screen "C5_GraphicView_2" 1024x768, template "T_C05"
   GraphicView "PNG_160x60_FitF" at 6,40 size 160x60; Picture "G_PNG"
   TextField "Label_PNG_160x60_FitF" at 6,102 size 113x20; Text 'PNG_160x60_FitF'
   GraphicView "PNG_160x60_FitT" at 182,40 size 160x60; Picture "G_PNG"
   TextField "Label_PNG_160x60_FitT" at 182,102 size 114x20; Text 'PNG_160x60_FitT'
   GraphicView "PNG_60x120_FitF" at 358,40 size 60x120; Picture "G_PNG"
   TextField "Label_PNG_60x120_FitF" at 358,162 size 113x20; Text 'PNG_60x120_FitF'
   GraphicView "PNG_60x120_FitT" at 534,40 size 60x120; Picture "G_PNG"
   TextField "Label_PNG_60x120_FitT" at 534,162 size 114x20; Text 'PNG_60x120_FitT'
   GraphicView "PNG_80x80_FitF" at 710,40 size 80x80; Picture "G_PNG"
   TextField "Label_PNG_80x80_FitF" at 710,122 size 105x20; Text 'PNG_80x80_FitF'
   GraphicView "PNG_80x80_FitT" at 6,182 size 80x80; Picture "G_PNG"
   TextField "Label_PNG_80x80_FitT" at 6,264 size 106x20; Text 'PNG_80x80_FitT'
   GraphicView "TALL_160x60_FitF" at 182,182 size 160x60; Picture "G_TALL"
   TextField "Label_TALL_160x60_FitF" at 182,244 size 120x20; Text 'TALL_160x60_FitF'
   GraphicView "TALL_160x60_FitT" at 358,182 size 160x60; Picture "G_TALL"
   TextField "Label_TALL_160x60_FitT" at 358,244 size 121x20; Text 'TALL_160x60_FitT'
   GraphicView "TALL_60x120_FitF" at 534,182 size 60x120; Picture "G_TALL"
   TextField "Label_TALL_60x120_FitF" at 534,304 size 120x20; Text 'TALL_60x120_FitF'
   GraphicView "TALL_60x120_FitT" at 710,182 size 60x120; Picture "G_TALL"
   TextField "Label_TALL_60x120_FitT" at 710,304 size 121x20; Text 'TALL_60x120_FitT'
   GraphicView "TALL_80x80_FitF" at 6,324 size 80x80; Picture "G_TALL"
   TextField "Label_TALL_80x80_FitF" at 6,406 size 112x20; Text 'TALL_80x80_FitF'
   GraphicView "TALL_80x80_FitT" at 182,324 size 80x80; Picture "G_TALL"
   TextField "Label_TALL_80x80_FitT" at 182,406 size 113x20; Text 'TALL_80x80_FitT'
   GraphicView "WIDE_160x60_FitF" at 358,324 size 160x60; Picture "G_WIDE"
   TextField "Label_WIDE_160x60_FitF" at 358,386 size 123x20; Text 'WIDE_160x60_FitF'
   GraphicView "WIDE_160x60_FitT" at 534,324 size 160x60; Picture "G_WIDE"
   TextField "Label_WIDE_160x60_FitT" at 534,386 size 124x20; Text 'WIDE_160x60_FitT'
   GraphicView "WIDE_60x120_FitF" at 710,324 size 60x120; Picture "G_WIDE"
   TextField "Label_WIDE_60x120_FitF" at 710,446 size 123x20; Text 'WIDE_60x120_FitF'
   GraphicView "WIDE_60x120_FitT" at 6,466 size 60x120; Picture "G_WIDE"
   TextField "Label_WIDE_60x120_FitT" at 6,588 size 124x20; Text 'WIDE_60x120_FitT'
   GraphicView "WIDE_80x80_FitF" at 182,466 size 80x80; Picture "G_WIDE"
   TextField "Label_WIDE_80x80_FitF" at 182,548 size 115x20; Text 'WIDE_80x80_FitF'
   GraphicView "WIDE_80x80_FitT" at 358,466 size 80x80; Picture "G_WIDE"
   TextField "Label_WIDE_80x80_FitT" at 358,548 size 116x20; Text 'WIDE_80x80_FitT'
   GraphicView "BMP_Transparent" at 534,466 size 120x80; Picture "G_BMP"
   TextField "Label_BMP_Transparent" at 534,548 size 120x20; Text 'BMP_Transparent'
   GraphicView "PNG_BackTransparent" at 710,466 size 120x80; Picture "G_PNG"
   TextField "Label_PNG_BackTransparent" at 710,548 size 147x20; Text 'PNG_BackTransparent'
   IOField "State" at 4,742 size 60x22; FormatPattern 9
      ProcessValue <- "D_State"
   Button "S1" at 70,742 size 40x22; TextOff 'S1'
      on Click: "SetS1"()
   Button "S2" at 114,742 size 40x22; TextOff 'S2'
      on Click: "SetS2"()
   Button "S3" at 158,742 size 40x22; TextOff 'S3'
      on Click: "SetS3"()
   Button "S4" at 202,742 size 40x22; TextOff 'S4'
      on Click: "SetS4"()
   Button "Next" at 980,742 size 40x22; TextOff 'Next'
      on Click: ActivateScreen("C5_Lists", 0)

screen "C5_Lists" 1024x768, template "T_C05"
   SymbolicIOField "SIO_TL_Value" at 6,40 size 160x30; TextOff '0'; TextOn '1'; TextList "TL_Value"
      ProcessValue <- "D_TL"
   TextField "Label_SIO_TL_Value" at 6,72 size 93x20; Text 'SIO_TL_Value'
   SymbolicIOField "SIO_TL_Bit" at 182,40 size 160x30; TextOff '0'; TextOn '1'; TextList "TL_Bit"
      ProcessValue <- "D_Bool"
   TextField "Label_SIO_TL_Bit" at 182,72 size 74x20; Text 'SIO_TL_Bit'
   SymbolicIOField "SIO_TL_BitNo" at 358,40 size 160x30; TextOff '0'; TextOn '1'; TextList "TL_BitNo"
      ProcessValue <- "D_Bits"
   TextField "Label_SIO_TL_BitNo" at 358,72 size 90x20; Text 'SIO_TL_BitNo'
   SymbolicIOField "SIO_TL_Value_Out" at 534,40 size 160x30; TextOff '0'; TextOn '1'; TextList "TL_Value"
      ProcessValue <- "D_TL"
   TextField "Label_SIO_TL_Value_Out" at 534,72 size 124x20; Text 'SIO_TL_Value_Out'
   GraphicIOField "GIO_GL_Value" at 710,40 size 120x80; PictureList "GL_Value"
      ProcessValue <- "D_TL"
   TextField "Label_GIO_GL_Value" at 710,122 size 94x20; Text 'GIO_GL_Value'
   GraphicIOField "GIO_GL_Bit" at 6,142 size 120x80; PictureList "GL_Bit"
      ProcessValue <- "D_Bool"
   TextField "Label_GIO_GL_Bit" at 6,224 size 75x20; Text 'GIO_GL_Bit'
   GraphicIOField "GIO_GL_BitNo" at 182,142 size 120x80; PictureList "GL_BitNo"
      ProcessValue <- "D_Bits"
   TextField "Label_GIO_GL_BitNo" at 182,224 size 91x20; Text 'GIO_GL_BitNo'
   GraphicIOField "GIO_GL_Value_Out" at 358,142 size 120x80; PictureList "GL_Value"
      ProcessValue <- "D_TL"
   TextField "Label_GIO_GL_Value_Out" at 358,224 size 125x20; Text 'GIO_GL_Value_Out'
   IOField "State" at 4,742 size 60x22; FormatPattern 9
      ProcessValue <- "D_State"
   Button "S1" at 70,742 size 40x22; TextOff 'S1'
      on Click: "SetS1"()
   Button "S2" at 114,742 size 40x22; TextOff 'S2'
      on Click: "SetS2"()
   Button "S3" at 158,742 size 40x22; TextOff 'S3'
      on Click: "SetS3"()
   Button "S4" at 202,742 size 40x22; TextOff 'S4'
      on Click: "SetS4"()
   Button "Next" at 980,742 size 40x22; TextOff 'Next'
      on Click: ActivateScreen("C5_Buttons", 0)

Template "T_C05" 1024x768
   TextField "T_Title" at 8,6 size 185x21; Text 'Template T_C05 (header)'
   DateTimeField "T_Clock" at 834,4 size 189x26

PopupScreen "Popup_C05" 300x200
   TextField "Pop_Title" at 10,10 size 175x20; Text 'Pop-up screen Popup_C05'
   GraphicView "Pop_Graphic" at 10,40 size 120x80; Picture "G_PNG"
   IOField "Pop_Value" at 150,60 size 120x30; FormatPattern s99999
      ProcessValue <- "D_Int"
   Button "Pop_Close" at 200,160 size 80x22; TextOff 'Close'
      on Click: function_efd93a16("Popup_C05", 200, 120, -1, -1, 1)

screen "C5_Structure" 1024x768, template "T_C05"
   Group "Group_A" at 10,50 size 300x85
   TextField "Label_Group_A (contains Group_B)" at 10,140 size 190x20; Text 'Group_A (contains Group_B)'
   TextField "Layer0_Text" at 352,52 size 54x20; Text 'Layer 0'
   TextField "Label_Layers 0-3 (layer 2 VisibleES false)" at 350,200 size 231x20; Text 'Layers 0-3 (layer 2 VisibleES false)'
   IOField "State" at 4,742 size 60x22; FormatPattern 9
      ProcessValue <- "D_State"
   Button "S1" at 70,742 size 40x22; TextOff 'S1'
      on Click: "SetS1"()
   Button "S2" at 114,742 size 40x22; TextOff 'S2'
      on Click: "SetS2"()
   Button "S3" at 158,742 size 40x22; TextOff 'S3'
      on Click: "SetS3"()
   Button "S4" at 202,742 size 40x22; TextOff 'S4'
      on Click: "SetS4"()
   Button "Popup" at 246,742 size 60x22; TextOff 'Popup'
      on Click: function_efd93a16("Popup_C05", 200, 120, -1, -1, 1)
   Button "SlideIn" at 310,742 size 60x22; TextOff 'Slide'
      on Click: "C5_ToggleSlideIn"()
   Button "Next" at 980,742 size 40x22; TextOff 'Next'
      on Click: ActivateScreen("C5_GraphicView_1", 0)
   Group "Group_B" at 210,50 size 100x85
   TextField "GB_Text" at 210,115 size 59x20; Text 'Group_B'
   TextField "Layer1_Text" at 382,72 size 54x20; Text 'Layer 1'
   TextField "Layer2_Text" at 412,92 size 54x20; Text 'Layer 2'
   TextField "Layer3_Text" at 442,112 size 54x20; Text 'Layer 3'

screen "C6_Faceplates" 1024x768
   ScreenModuleView "FP_Dyn" at 10,10 size 300x150; ScreenModuleType ""; Guid_{11997190-83750} 'Tags D_Int D_Range D_Pct'
      Guid_{11997190-83886} <- "D_Int"
      Guid_{11997190-83896} <- "D_Range"
      Guid_{11997190-83898} <- "D_Pct"
      Guid_{11997190-83900} <- "D_Vis"
   TextField "Label_FP_Dyn" at 10,162 size 52x20; Text 'FP_Dyn'
   ScreenModuleView "FP_Static" at 330,10 size 300x150; ScreenModuleType ""; Guid_{11997190-83750} 'Static values'
   TextField "Label_FP_Static" at 330,162 size 65x20; Text 'FP_Static'
   ScreenModuleView "FP_Alt" at 10,186 size 300x150; ScreenModuleType ""; Guid_{11997190-83750} 'Tags D_SInt D_TL D_UInt'
      Guid_{11997190-83886} <- "D_SInt"
      Guid_{11997190-83896} <- "D_TL"
      Guid_{11997190-83898} <- "D_UInt"
      Guid_{11997190-83900} <- "D_En"
   TextField "Label_FP_Alt" at 10,338 size 46x20; Text 'FP_Alt'
   ScreenModuleView "FP_Move" at 330,186 size 300x150; ScreenModuleType ""; Guid_{11997190-83750} 'Moved by D_Pct'
      Guid_{11997190-83886} <- "D_Int"
      Guid_{11997190-83896} <- "D_Range"
      Guid_{11997190-83898} <- "D_Pct"
      Guid_{11997190-83900} <- "D_Vis"
      HorizontalMovement <- "D_Pct"
   TextField "Label_FP_Move" at 330,338 size 62x20; Text 'FP_Move'
   IOField "State" at 4,742 size 60x22; FormatPattern 9
      ProcessValue <- "D_State"
   Button "S1" at 70,742 size 40x22; TextOff 'S1'
      on Click: "SetS1"()
   Button "S2" at 114,742 size 40x22; TextOff 'S2'
      on Click: "SetS2"()
   Button "S3" at 158,742 size 40x22; TextOff 'S3'
      on Click: "SetS3"()
   Button "S4" at 202,742 size 40x22; TextOff 'S4'
      on Click: "SetS4"()
   Button "Next" at 980,742 size 40x22; TextOff 'Next'
      on Click: ActivateScreen("C6_Faceplates", 0)

VB script "C5_ToggleSlideIn"
   ' slide-in screens are not available on WinCC RT Advanced

VB script "SetS1"
   SmartTags("D_State") = 1
   SmartTags("D_Bool") = False
   SmartTags("D_SInt") = -128
   SmartTags("D_Int") = -32768
   SmartTags("D_DInt") = -2147483648
   SmartTags("D_USInt") = 0
   SmartTags("D_UInt") = 0
   SmartTags("D_UDInt") = 0
   SmartTags("D_Real") = -999.999
   SmartTags("D_LReal") = -0.00000015
   SmartTags("D_String") = ""
   SmartTags("D_DateTime") = DateSerial(1990, 1, 1) + TimeSerial(0, 0, 0)
   SmartTags("D_Pct") = 0
   SmartTags("D_Range") = 5
   SmartTags("D_Bits") = 1
   SmartTags("D_Vis") = False
   SmartTags("D_En") = False
   SmartTags("D_X") = 10
   SmartTags("D_Y") = 10
   SmartTags("D_Max") = 100
   SmartTags("D_Min") = 0
   SmartTags("D_TL") = -5
   SmartTags("D_BarR") = -5

VB script "SetS2"
   SmartTags("D_State") = 2
   SmartTags("D_Bool") = True
   SmartTags("D_SInt") = 12
   SmartTags("D_Int") = 1234
   SmartTags("D_DInt") = 123456
   SmartTags("D_USInt") = 200
   SmartTags("D_UInt") = 40000
   SmartTags("D_UDInt") = 3000000000
   SmartTags("D_Real") = 3.14159
   SmartTags("D_LReal") = 2.718281828
   SmartTags("D_String") = "Hello World"
   SmartTags("D_DateTime") = DateSerial(2026, 11, 22) + TimeSerial(13, 45, 30)
   SmartTags("D_Pct") = 50
   SmartTags("D_Range") = 25
   SmartTags("D_Bits") = 2
   SmartTags("D_Vis") = True
   SmartTags("D_En") = True
   SmartTags("D_X") = 256
   SmartTags("D_Y") = 192
   SmartTags("D_Max") = 200
   SmartTags("D_Min") = -100
   SmartTags("D_TL") = 5
   SmartTags("D_BarR") = 0

VB script "SetS3"
   SmartTags("D_State") = 3
   SmartTags("D_Bool") = True
   SmartTags("D_SInt") = 127
   SmartTags("D_Int") = 32767
   SmartTags("D_DInt") = 2147483647
   SmartTags("D_USInt") = 255
   SmartTags("D_UInt") = 65535
   SmartTags("D_UDInt") = 4294967295
   SmartTags("D_Real") = 123456.789
   SmartTags("D_LReal") = 1E+300
   SmartTags("D_String") = "Ünïcödé äöüß ÄÖÜ € – long text that is wider than the field 0123456789 ABCDEFGHIJ"
   SmartTags("D_DateTime") = DateSerial(2099, 12, 31) + TimeSerial(23, 59, 59)
   SmartTags("D_Pct") = 100
   SmartTags("D_Range") = 75
   SmartTags("D_Bits") = 4
   SmartTags("D_Vis") = True
   SmartTags("D_En") = False
   SmartTags("D_X") = 682
   SmartTags("D_Y") = 384
   SmartTags("D_Max") = 50
   SmartTags("D_Min") = -50
   SmartTags("D_TL") = 10
   SmartTags("D_BarR") = 5

VB script "SetS4"
   SmartTags("D_State") = 4
   SmartTags("D_Bool") = False
   SmartTags("D_SInt") = -1
   SmartTags("D_Int") = -1
   SmartTags("D_DInt") = 0
   SmartTags("D_USInt") = 1
   SmartTags("D_UInt") = 1
   SmartTags("D_UDInt") = 1
   SmartTags("D_Real") = 0.0005
   SmartTags("D_LReal") = -0.0
   SmartTags("D_String") = "äöü ÄÖÜ ß"
   SmartTags("D_DateTime") = DateSerial(1970, 1, 1) + TimeSerial(0, 0, 0)
   SmartTags("D_Pct") = 150
   SmartTags("D_Range") = 200
   SmartTags("D_Bits") = 9
   SmartTags("D_Vis") = False
   SmartTags("D_En") = True
   SmartTags("D_X") = -20
   SmartTags("D_Y") = 0
   SmartTags("D_Max") = 100
   SmartTags("D_Min") = 0
   SmartTags("D_TL") = 50
   SmartTags("D_BarR") = 2.5
*)

(* ===== HMI "HMI_TP900S" =====
system functions are stored by id; their names below are inferred from use

HMI tags "Default tag table"
   "Hmi_Bool" : Bool, internal
   "Hmi_Int" : Int, internal
   "Hmi_Real" : Real, internal
   "Hmi_String" : WString[254], internal

screen "All_Objects" 800x480
   TextField "TextField_1" at 680,10 size 35x17; Text 'Text'
   GraphicView "GraphicView_1" at 10,80 size 100x60
   IOField "IOField_1" at 130,80 size 100x30
   Button "Button_1" at 250,80 size 100x40; TextOff 'Text'
   SymbolicIOField "SymbolicIOField_1" at 370,80 size 120x30; TextOff '0'; TextOn '1'
   GraphicIOField "GraphicIOField_1" at 510,80 size 60x60
   DateTimeField "DateTimeField_1" at 590,80 size 189x26
   Bar "Bar_1" at 10,160 size 40x120
   Switch "Switch_1" at 70,160 size 120x40; CaptionText 'Switch'; TextOff '0'; TextOn '1'
   SymbolLibrary "SymbolLibrary_1" at 210,160 size 60x60
   Slider "Slider_1" at 290,160 size 60x160; Caption 'SIMATIC'
   Gauge "Gauge_1" at 370,160 size 150x150; CaptionText 'SIMATIC'
   Clock "Clock_1" at 540,160 size 150x150

screen "Ctl_01_AlarmView" 800x480, template "Nav"
   AlarmView "Alarm view_1" at 3,3 size 600x300

screen "Ctl_02_TrendView" 800x480, template "Nav"
   TrendView "Trend view_1" at 3,3 size 600x300

screen "Ctl_03_UserView" 800x480, template "Nav"
   UserView "User view_1" at 3,3 size 480x240

screen "Ctl_04_HtmlBrowser" 800x480, template "Nav"
   HTMLBrowser "HTML browser_1" at 3,3 size 192x192

screen "Ctl_05_WatchTable" 800x480, template "Nav"
   StatusForce "Watch table_1" at 3,3 size 600x300; ToolTipText 'Text'

screen "Ctl_06_SmartClientView" 800x480, template "Nav"
   SmartClientView "Sm@rtClient view_1" at 3,3 size 320x240

screen "Ctl_07_RecipeView" 800x480, template "Nav"
   RecipeView "Recipe view_1" at 3,3 size 400x330

screen "Ctl_09_SysDiagView" 800x480, template "Nav"
   SysDiagControl "System diagnostics view_1" at 3,3 size 600x300

screen "Ctl_10_MediaPlayer" 800x480, template "Nav"
   MediaPlayer "Media Player_1" at 3,3 size 240x240

screen "Ctl_11_PlcCodeView" 800x480, template "Nav"
   PLCCodeViewer "PLC code view_1" at 3,3 size 600x300

screen "Ctl_12_GraphOverview" 800x480, template "Nav"
   S7GraphOverview "GRAPH overview_1" at 3,3 size 424x72

screen "Ctl_13_ProDiagOverview" 800x480, template "Nav"
   ProDiagOverview "ProDiag overview_1" at 3,3 size 253x72

screen "Ctl_14_CriteriaAnalysisView" 800x480, template "Nav"
   CriteriaAnalysisView "Criteria analysis view_1" at 3,3 size 460x150

screen "Ctl_15_CameraView" 800x480, template "Nav"
   CameraControl "Camera view_1" at 3,3 size 320x240

screen "Ctl_16_PdfView" 800x480, template "Nav"
   PDFView "PDFView_1" at 3,3 size 320x240

Template "Nav" 800x480
   Button "Nav_01" at 770,2 size 28x22; TextOff 'Text'
      on Click: ActivateScreen("Ctl_01_AlarmView", 0)
   Button "Nav_02" at 770,28 size 28x22; TextOff 'Text'
      on Click: ActivateScreen("Ctl_02_TrendView", 0)
   Button "Nav_03" at 770,54 size 28x22; TextOff 'Text'
      on Click: ActivateScreen("Ctl_03_UserView", 0)
   Button "Nav_04" at 770,80 size 28x22; TextOff 'Text'
      on Click: ActivateScreen("Ctl_04_HtmlBrowser", 0)
   Button "Nav_05" at 770,106 size 28x22; TextOff 'Text'
      on Click: ActivateScreen("Ctl_05_WatchTable", 0)
   Button "Nav_06" at 770,132 size 28x22; TextOff 'Text'
      on Click: ActivateScreen("Ctl_06_SmartClientView", 0)
   Button "Nav_07" at 770,158 size 28x22; TextOff 'Text'
      on Click: ActivateScreen("Ctl_07_RecipeView", 0)
   Button "Nav_09" at 770,210 size 28x22; TextOff 'Text'
      on Click: ActivateScreen("Ctl_09_SysDiagView", 0)
   Button "Nav_10" at 770,236 size 28x22; TextOff 'Text'
      on Click: ActivateScreen("Ctl_10_MediaPlayer", 0)
   Button "Nav_11" at 770,262 size 28x22; TextOff 'Text'
      on Click: ActivateScreen("Ctl_11_PlcCodeView", 0)
   Button "Nav_12" at 770,288 size 28x22; TextOff 'Text'
      on Click: ActivateScreen("Ctl_12_GraphOverview", 0)
   Button "Nav_13" at 770,314 size 28x22; TextOff 'Text'
      on Click: ActivateScreen("Ctl_13_ProDiagOverview", 0)
   Button "Nav_14" at 770,340 size 28x22; TextOff 'Text'
      on Click: ActivateScreen("Ctl_14_CriteriaAnalysisView", 0)
   Button "Nav_15" at 770,366 size 28x22; TextOff 'Text'
      on Click: ActivateScreen("Ctl_15_CameraView", 0)
   Button "Nav_16" at 770,392 size 28x22; TextOff 'Text'
      on Click: ActivateScreen("Ctl_16_PdfView", 0)
   Button "Nav_17" at 770,418 size 28x22; TextOff 'Text'
      on Click: ActivateScreen("All_Objects", 0)
*)

(* ===== HMI "HMI_TP1200" =====
system functions are stored by id; their names below are inferred from use
connection "HMI_Connection_4": ETHERNET, S7_1500_OMS

HMI tags "Default tag table"
   "Hmi_Bool" : Bool, internal
   "Hmi_Int" : Int, internal
   "Hmi_Real" : Real, internal
   "Hmi_String" : WString[254], internal
   "Ext_Bool" : Bool = PLC Plc_Bool AT %M100.0, 1 s
   "Ext_Int" : Int = PLC Plc_Int AT %MW102, 1 s
   "Ext_Real" : Real = PLC Plc_Real AT %MD104, 1 s
   "Ext_Byte" : Byte = PLC Plc_Byte AT %MB108, 1 s

HMI tags "C03_Tags"
   "D_State" : Int, internal
   "D_Bool" : Bool, internal
   "D_SInt" : SInt, internal
   "D_Int" : Int, internal
   "D_DInt" : DInt, internal
   "D_USInt" : USInt, internal
   "D_UInt" : UInt, internal
   "D_UDInt" : UDInt, internal
   "D_Real" : Real, internal
   "D_LReal" : LReal, internal
   "D_String" : WString[254], internal
   "D_DateTime" : DateTime, internal
   "D_Pct" : Int, internal
   "D_Range" : Int, internal
   "D_Bits" : Int, internal
   "D_Vis" : Bool, internal
   "D_En" : Bool, internal
   "D_X" : Int, internal
   "D_Y" : Int, internal
   "D_Max" : Real, internal
   "D_Min" : Real, internal
   "D_TL" : Int, internal
   "D_BarR" : Real, internal

discrete alarms
   1: 'Alarm bit 0 (D_Bits)', class Errors, trigger "D_Bits" bit 0
   2: 'Alarm bit 1 (D_Bits)', class Errors, trigger "D_Bits" bit 1
   3: 'Alarm bit 2 (D_Bits)', class Warnings, trigger "D_Bits" bit 2
   4: 'Alarm bit 3 (D_Bits)', class Warnings, trigger "D_Bits" bit 3

analog alarms
   1: 'D_Range above 50', class Errors, trigger "D_Range"

text list "TL_Bit": 0 'Off (0)'; 1 'On (1)'

text list "TL_BitNo": 0 'Bit 0 set'; 1 'Bit 1 set'; 2 'Bit 2 set'; 3 'Bit 3 set'

text list "TL_Value": -100..-1 'Negative (-100..-1)'; 0 'Zero'; 1..9 'One to nine'; 10 'Ten: Ünïcödé äöüß ÄÖÜ €'; 32000 'Undefined value (default entry)'

graphic list "GL_Bit": 0 'G_EMF'; 1 'G_WMF'

graphic list "GL_BitNo": 0 'G_PNG'; 1 'G_JPG'; 2 'G_BMP'; 3 'G_TIF'

graphic list "GL_Value": -100..-1 'G_GIF'; 0 'G_PNG'; 1..9 'G_JPG'; 10 'G_BMP'; 32000 'G_SVG'

recipe "Recipe_1": Recipe_element_1 <- "D_Int", Recipe_element_2 <- "D_Real", Recipe_element_3 <- "D_Pct", Recipe_element_4 <- "D_Bits", Recipe_element_5 <- "D_Range"

SlideinScreen "GraphX_Slidein_Top" 1280x120
   TextField "SI_Title" at 10,10 size 167x22; Text 'Slide-in screen Top'
   Bar "SI_Bar" at 330,10 size 200x40
      ProcessValue <- "D_Pct"
   IOField "SI_Value" at 560,10 size 120x30; FormatPattern s99999
      ProcessValue <- "D_Int"

screen "All_Objects" 1280x800
   TextField "TextField_1" at 680,10 size 42x22; Text 'Text'
   GraphicView "GraphicView_1" at 800,10 size 100x60
   IOField "IOField_1" at 920,10 size 100x30
   Button "Button_1" at 1040,10 size 100x40; TextOff 'Text'
   SymbolicIOField "SymbolicIOField_1" at 10,90 size 120x30; TextOff '0'; TextOn '1'
   GraphicIOField "GraphicIOField_1" at 150,90 size 60x60
   DateTimeField "DateTimeField_1" at 230,90 size 189x26
   Bar "Bar_1" at 410,90 size 40x120
   Switch "Switch_1" at 470,90 size 120x40; CaptionText 'Switch'; TextOff '0'; TextOn '1'
   SymbolLibrary "SymbolLibrary_1" at 610,90 size 60x60
   Slider "Slider_1" at 690,90 size 60x160; Caption 'SIMATIC'
   Gauge "Gauge_1" at 770,90 size 150x150; CaptionText 'SIMATIC'
   Clock "Clock_1" at 940,90 size 150x150

screen "Ctl_01_AlarmView" 1280x800, template "Nav"
   AlarmView "Alarm view_1" at 3,3 size 600x300

screen "Ctl_02_TrendView" 1280x800, template "Nav"
   TrendView "Trend view_1" at 3,3 size 600x300

screen "Ctl_03_UserView" 1280x800, template "Nav"
   UserView "User view_1" at 3,3 size 480x240

screen "Ctl_04_HtmlBrowser" 1280x800, template "Nav"
   HTMLBrowser "HTML browser_1" at 3,3 size 192x192

screen "Ctl_05_WatchTable" 1280x800, template "Nav"
   StatusForce "Watch table_1" at 3,3 size 600x300; ToolTipText 'Text'

screen "Ctl_06_SmartClientView" 1280x800, template "Nav"
   SmartClientView "Sm@rtClient view_1" at 3,3 size 320x240

screen "Ctl_07_RecipeView" 1280x800, template "Nav"
   RecipeView "Recipe view_1" at 3,3 size 400x330; Recipe "Recipe_1"

screen "Ctl_09_SysDiagView" 1280x800, template "Nav"
   SysDiagControl "System diagnostics view_1" at 3,3 size 600x300

screen "Ctl_10_MediaPlayer" 1280x800, template "Nav"
   MediaPlayer "Media Player_1" at 3,3 size 240x240

screen "Ctl_15_CameraView" 1280x800, template "Nav"
   CameraControl "Camera view_1" at 3,3 size 320x240

screen "Ctl_16_PdfView" 1280x800, template "Nav"
   PDFView "PDFView_1" at 3,3 size 320x240

Template "Nav" 1280x800
   Button "Nav_01" at 1250,2 size 28x22; TextOff 'Text'
      on Click: ActivateScreen("Ctl_01_AlarmView", 0)
   Button "Nav_02" at 1250,28 size 28x22; TextOff 'Text'
      on Click: ActivateScreen("Ctl_02_TrendView", 0)
   Button "Nav_03" at 1250,54 size 28x22; TextOff 'Text'
      on Click: ActivateScreen("Ctl_03_UserView", 0)
   Button "Nav_04" at 1250,80 size 28x22; TextOff 'Text'
      on Click: ActivateScreen("Ctl_04_HtmlBrowser", 0)
   Button "Nav_05" at 1250,106 size 28x22; TextOff 'Text'
      on Click: ActivateScreen("Ctl_05_WatchTable", 0)
   Button "Nav_06" at 1250,132 size 28x22; TextOff 'Text'
      on Click: ActivateScreen("Ctl_06_SmartClientView", 0)
   Button "Nav_07" at 1250,158 size 28x22; TextOff 'Text'
      on Click: ActivateScreen("Ctl_07_RecipeView", 0)
   Button "Nav_09" at 1250,210 size 28x22; TextOff 'Text'
      on Click: ActivateScreen("Ctl_09_SysDiagView", 0)
   Button "Nav_10" at 1250,236 size 28x22; TextOff 'Text'
      on Click: ActivateScreen("Ctl_10_MediaPlayer", 0)
   Button "Nav_15" at 1250,366 size 28x22; TextOff 'Text'
      on Click: ActivateScreen("Ctl_15_CameraView", 0)
   Button "Nav_16" at 1250,392 size 28x22; TextOff 'Text'
      on Click: ActivateScreen("Ctl_16_PdfView", 0)
   Button "Nav_17" at 1250,418 size 28x22; TextOff 'Text'
      on Click: ActivateScreen("All_Objects", 0)

screen "P_Line_1" 1280x800
   TextField "Label_Default" at 10,62 size 67x22; Text 'Default'
   TextField "Label_BackColor" at 120,62 size 90x22; Text 'BackColor'
   TextField "Label_Color" at 230,62 size 50x22; Text 'Color'
   TextField "Label_EndStyle" at 340,62 size 79x22; Text 'EndStyle'
   TextField "Label_EndStyle_2" at 450,62 size 101x22; Text 'EndStyle_2'
   TextField "Label_EndStyle_3" at 560,62 size 101x22; Text 'EndStyle_3'
   TextField "Label_EndStyle_4" at 670,62 size 101x22; Text 'EndStyle_4'
   TextField "Label_EndStyle_5" at 780,62 size 101x22; Text 'EndStyle_5'
   TextField "Label_FillStyle" at 890,62 size 77x22; Text 'FillStyle'
   TextField "Label_Flashing" at 1000,62 size 76x22; Text 'Flashing'
   TextField "Label_LineEndShapeStyle_2" at 1110,62 size 188x22; Text 'LineEndShapeStyle_2'
   TextField "Label_LineWidth" at 10,138 size 90x22; Text 'LineWidth'
   TextField "Label_StartStyle" at 120,138 size 92x22; Text 'StartStyle'
   TextField "Label_StartStyle_2" at 230,138 size 114x22; Text 'StartStyle_2'
   TextField "Label_StartStyle_3" at 340,138 size 114x22; Text 'StartStyle_3'
   TextField "Label_StartStyle_4" at 450,138 size 114x22; Text 'StartStyle_4'
   TextField "Label_StartStyle_5" at 560,138 size 114x22; Text 'StartStyle_5'
   TextField "Label_Style" at 670,138 size 49x22; Text 'Style'
   TextField "Label_Style_2" at 780,138 size 71x22; Text 'Style_2'
   TextField "Label_Style_3" at 890,138 size 71x22; Text 'Style_3'
   TextField "Label_Style_4" at 1000,138 size 71x22; Text 'Style_4'
   TextField "Label_UseDesignColorSchema" at 1110,138 size 202x22; Text 'UseDesignColorSchema'
   Button "Next" at 1238,776 size 40x22; TextOff 'Text'
      on Click: ActivateScreen("P_Polyline_1", 0)

screen "P_Polyline_1" 1280x800
   TextField "Label_Default" at 10,62 size 67x22; Text 'Default'
   TextField "Label_BackColor" at 120,62 size 90x22; Text 'BackColor'
   TextField "Label_Color" at 230,62 size 50x22; Text 'Color'
   TextField "Label_EndStyle" at 340,62 size 79x22; Text 'EndStyle'
   TextField "Label_EndStyle_2" at 450,62 size 101x22; Text 'EndStyle_2'
   TextField "Label_EndStyle_3" at 560,62 size 101x22; Text 'EndStyle_3'
   TextField "Label_EndStyle_4" at 670,62 size 101x22; Text 'EndStyle_4'
   TextField "Label_EndStyle_5" at 780,62 size 101x22; Text 'EndStyle_5'
   TextField "Label_FillStyle" at 890,62 size 77x22; Text 'FillStyle'
   TextField "Label_Flashing" at 1000,62 size 76x22; Text 'Flashing'
   TextField "Label_LineEndShapeStyle_2" at 1110,62 size 188x22; Text 'LineEndShapeStyle_2'
   TextField "Label_LineWidth" at 10,138 size 90x22; Text 'LineWidth'
   TextField "Label_StartStyle" at 120,138 size 92x22; Text 'StartStyle'
   TextField "Label_StartStyle_2" at 230,138 size 114x22; Text 'StartStyle_2'
   TextField "Label_StartStyle_3" at 340,138 size 114x22; Text 'StartStyle_3'
   TextField "Label_StartStyle_4" at 450,138 size 114x22; Text 'StartStyle_4'
   TextField "Label_StartStyle_5" at 560,138 size 114x22; Text 'StartStyle_5'
   TextField "Label_Style" at 670,138 size 49x22; Text 'Style'
   TextField "Label_Style_2" at 780,138 size 71x22; Text 'Style_2'
   TextField "Label_Style_3" at 890,138 size 71x22; Text 'Style_3'
   TextField "Label_Style_4" at 1000,138 size 71x22; Text 'Style_4'
   TextField "Label_UseDesignColorSchema" at 1110,138 size 202x22; Text 'UseDesignColorSchema'
   Button "Next" at 1238,776 size 40x22; TextOff 'Text'
      on Click: ActivateScreen("P_Polygon_1", 0)

screen "P_Polygon_1" 1280x800
   TextField "Label_Default" at 10,62 size 67x22; Text 'Default'
   TextField "Label_BackColor" at 120,62 size 90x22; Text 'BackColor'
   TextField "Label_BackFillStyle" at 230,62 size 117x22; Text 'BackFillStyle'
   TextField "Label_BorderColor" at 340,62 size 107x22; Text 'BorderColor'
   TextField "Label_BorderWidth" at 450,62 size 111x22; Text 'BorderWidth'
   TextField "Label_EdgeStyle" at 560,62 size 89x22; Text 'EdgeStyle'
   TextField "Label_EdgeStyle_2" at 670,62 size 111x22; Text 'EdgeStyle_2'
   TextField "Label_EdgeStyle_3" at 780,62 size 111x22; Text 'EdgeStyle_3'
   TextField "Label_EdgeStyle_4" at 890,62 size 111x22; Text 'EdgeStyle_4'
   TextField "Label_Flashing" at 1000,62 size 76x22; Text 'Flashing'
   TextField "Label_UseDesignColorSchema" at 1110,62 size 202x22; Text 'UseDesignColorSchema'
   Button "Next" at 1238,776 size 40x22; TextOff 'Text'
      on Click: ActivateScreen("P_Ellipse_1", 0)

screen "P_Ellipse_1" 1280x800
   TextField "Label_Default" at 10,62 size 67x22; Text 'Default'
   TextField "Label_BackColor" at 120,62 size 90x22; Text 'BackColor'
   TextField "Label_BackFillStyle" at 230,62 size 117x22; Text 'BackFillStyle'
   TextField "Label_BorderColor" at 340,62 size 107x22; Text 'BorderColor'
   TextField "Label_BorderWidth" at 450,62 size 111x22; Text 'BorderWidth'
   TextField "Label_EdgeStyle" at 560,62 size 89x22; Text 'EdgeStyle'
   TextField "Label_EdgeStyle_2" at 670,62 size 111x22; Text 'EdgeStyle_2'
   TextField "Label_EdgeStyle_3" at 780,62 size 111x22; Text 'EdgeStyle_3'
   TextField "Label_EdgeStyle_4" at 890,62 size 111x22; Text 'EdgeStyle_4'
   TextField "Label_Flashing" at 1000,62 size 76x22; Text 'Flashing'
   TextField "Label_UseDesignColorSchema" at 1110,62 size 202x22; Text 'UseDesignColorSchema'
   Button "Next" at 1238,776 size 40x22; TextOff 'Text'
      on Click: ActivateScreen("P_Circle_1", 0)

screen "P_Circle_1" 1280x800
   TextField "Label_Default" at 10,62 size 67x22; Text 'Default'
   TextField "Label_BackColor" at 70,62 size 90x22; Text 'BackColor'
   TextField "Label_BackFillStyle" at 130,62 size 117x22; Text 'BackFillStyle'
   TextField "Label_BorderColor" at 190,62 size 107x22; Text 'BorderColor'
   TextField "Label_BorderWidth" at 250,62 size 111x22; Text 'BorderWidth'
   TextField "Label_EdgeStyle" at 310,62 size 89x22; Text 'EdgeStyle'
   TextField "Label_EdgeStyle_2" at 370,62 size 111x22; Text 'EdgeStyle_2'
   TextField "Label_EdgeStyle_3" at 430,62 size 111x22; Text 'EdgeStyle_3'
   TextField "Label_EdgeStyle_4" at 490,62 size 111x22; Text 'EdgeStyle_4'
   TextField "Label_Flashing" at 550,62 size 76x22; Text 'Flashing'
   TextField "Label_UseDesignColorSchema" at 610,62 size 202x22; Text 'UseDesignColorSchema'
   Button "Next" at 1238,776 size 40x22; TextOff 'Text'
      on Click: ActivateScreen("P_Rectangle_1", 0)

screen "P_Rectangle_1" 1280x800
   TextField "Label_Default" at 10,62 size 67x22; Text 'Default'
   TextField "Label_BackColor" at 120,62 size 90x22; Text 'BackColor'
   TextField "Label_BackFillStyle" at 230,62 size 117x22; Text 'BackFillStyle'
   TextField "Label_BorderColor" at 340,62 size 107x22; Text 'BorderColor'
   TextField "Label_BorderWidth" at 450,62 size 111x22; Text 'BorderWidth'
   TextField "Label_EdgeStyle" at 560,62 size 89x22; Text 'EdgeStyle'
   TextField "Label_EdgeStyle_2" at 670,62 size 111x22; Text 'EdgeStyle_2'
   TextField "Label_EdgeStyle_3" at 780,62 size 111x22; Text 'EdgeStyle_3'
   TextField "Label_EdgeStyle_4" at 890,62 size 111x22; Text 'EdgeStyle_4'
   TextField "Label_Flashing" at 1000,62 size 76x22; Text 'Flashing'
   TextField "Label_RoundCornerHeight" at 1110,62 size 169x22; Text 'RoundCornerHeight'
   TextField "Label_RoundCornerWidth" at 10,138 size 163x22; Text 'RoundCornerWidth'
   TextField "Label_UseDesignColorSchema" at 120,138 size 202x22; Text 'UseDesignColorSchema'
   Button "Next" at 1238,776 size 40x22; TextOff 'Text'
      on Click: ActivateScreen("P_TextField_1", 0)

screen "P_TextField_1" 1280x800
   TextField "Default" at 10,10 size 42x22; Text 'Text'
   TextField "Label_Default" at 10,42 size 67x22; Text 'Default'
   TextField "BackColor" at 120,10 size 42x22; Text 'Text'
   TextField "Label_BackColor" at 120,42 size 90x22; Text 'BackColor'
   TextField "BackFillStyle" at 230,10 size 42x22; Text 'Text'
   TextField "Label_BackFillStyle" at 230,42 size 117x22; Text 'BackFillStyle'
   TextField "BorderBackColor" at 340,10 size 42x22; Text 'Text'
   TextField "Label_BorderBackColor" at 340,42 size 147x22; Text 'BorderBackColor'
   TextField "BorderColor" at 450,10 size 42x22; Text 'Text'
   TextField "Label_BorderColor" at 450,42 size 107x22; Text 'BorderColor'
   TextField "BorderWidth" at 560,10 size 42x22; Text 'Text'
   TextField "Label_BorderWidth" at 560,42 size 111x22; Text 'BorderWidth'
   TextField "BottomMargin" at 670,10 size 42x22; Text 'Text'
   TextField "Label_BottomMargin" at 670,42 size 122x22; Text 'BottomMargin'
   TextField "CornerRadius" at 780,10 size 42x22; Text 'Text'
   TextField "Label_CornerRadius" at 780,42 size 119x22; Text 'CornerRadius'
   TextField "EdgeStyle" at 890,10 size 42x22; Text 'Text'
   TextField "Label_EdgeStyle" at 890,42 size 89x22; Text 'EdgeStyle'
   TextField "EdgeStyle_2" at 1000,10 size 42x22; Text 'Text'
   TextField "Label_EdgeStyle_2" at 1000,42 size 111x22; Text 'EdgeStyle_2'
   TextField "EdgeStyle_3" at 1110,10 size 42x22; Text 'Text'
   TextField "Label_EdgeStyle_3" at 1110,42 size 111x22; Text 'EdgeStyle_3'
   TextField "EdgeStyle_4" at 10,66 size 42x22; Text 'Text'
   TextField "Label_EdgeStyle_4" at 10,98 size 111x22; Text 'EdgeStyle_4'
   TextField "FitToLargest" at 120,66 size 100x30; Text 'Text'
   TextField "Label_FitToLargest" at 120,98 size 112x22; Text 'FitToLargest'
   TextField "Flashing" at 230,66 size 42x22; Text 'Text'
   TextField "Label_Flashing" at 230,98 size 76x22; Text 'Flashing'
   TextField "ForeColor" at 340,66 size 42x22; Text 'Text'
   TextField "Label_ForeColor" at 340,98 size 88x22; Text 'ForeColor'
   TextField "HorizontalAlignment" at 450,66 size 42x22; Text 'Text'
   TextField "Label_HorizontalAlignment" at 450,98 size 177x22; Text 'HorizontalAlignment'
   TextField "HorizontalAlignment_2" at 560,66 size 42x22; Text 'Text'
   TextField "Label_HorizontalAlignment_2" at 560,98 size 199x22; Text 'HorizontalAlignment_2'
   TextField "LeftMargin" at 670,66 size 42x22; Text 'Text'
   TextField "Label_LeftMargin" at 670,98 size 97x22; Text 'LeftMargin'
   TextField "RightMargin" at 780,66 size 42x22; Text 'Text'
   TextField "Label_RightMargin" at 780,98 size 108x22; Text 'RightMargin'
   TextField "TopMargin" at 890,66 size 42x22; Text 'Text'
   TextField "Label_TopMargin" at 890,98 size 93x22; Text 'TopMargin'
   TextField "UseDesignColorSchema" at 1000,66 size 33x21; Text 'Text'
   TextField "Label_UseDesignColorSchema" at 1000,98 size 202x22; Text 'UseDesignColorSchema'
   TextField "VerticalAlignment" at 1110,66 size 42x22; Text 'Text'
   TextField "Label_VerticalAlignment" at 1110,98 size 156x22; Text 'VerticalAlignment'
   TextField "VerticalAlignment_2" at 10,122 size 42x22; Text 'Text'
   TextField "Label_VerticalAlignment_2" at 10,154 size 178x22; Text 'VerticalAlignment_2'
   Button "Next" at 1238,776 size 40x22; TextOff 'Text'
      on Click: ActivateScreen("P_GraphicView_1", 0)

screen "P_GraphicView_1" 1280x800
   GraphicView "Default" at 10,10 size 100x60
   TextField "Label_Default" at 10,72 size 67x22; Text 'Default'
   GraphicView "BackColor" at 120,10 size 100x60
   TextField "Label_BackColor" at 120,72 size 90x22; Text 'BackColor'
   GraphicView "BackFillStyle" at 230,10 size 100x60
   TextField "Label_BackFillStyle" at 230,72 size 117x22; Text 'BackFillStyle'
   GraphicView "BorderColor" at 340,10 size 100x60
   TextField "Label_BorderColor" at 340,72 size 107x22; Text 'BorderColor'
   GraphicView "BorderWidth" at 450,10 size 100x60
   TextField "Label_BorderWidth" at 450,72 size 111x22; Text 'BorderWidth'
   GraphicView "EdgeStyle" at 560,10 size 100x60
   TextField "Label_EdgeStyle" at 560,72 size 89x22; Text 'EdgeStyle'
   GraphicView "EdgeStyle_2" at 670,10 size 100x60
   TextField "Label_EdgeStyle_2" at 670,72 size 111x22; Text 'EdgeStyle_2'
   GraphicView "EdgeStyle_3" at 780,10 size 100x60
   TextField "Label_EdgeStyle_3" at 780,72 size 111x22; Text 'EdgeStyle_3'
   GraphicView "EdgeStyle_4" at 890,10 size 100x60
   TextField "Label_EdgeStyle_4" at 890,72 size 111x22; Text 'EdgeStyle_4'
   GraphicView "FitToLargest" at 1000,10 size 100x60
   TextField "Label_FitToLargest" at 1000,72 size 112x22; Text 'FitToLargest'
   GraphicView "Flashing" at 1110,10 size 100x60
   TextField "Label_Flashing" at 1110,72 size 76x22; Text 'Flashing'
   GraphicView "TransparentColor" at 10,96 size 100x60
   TextField "Label_TransparentColor" at 10,158 size 152x22; Text 'TransparentColor'
   GraphicView "UseTransparentColor" at 120,96 size 100x60
   TextField "Label_UseTransparentColor" at 120,158 size 183x22; Text 'UseTransparentColor'
   Button "Next" at 1238,776 size 40x22; TextOff 'Text'
      on Click: ActivateScreen("P_IOField_1", 0)

screen "P_IOField_1" 1280x800
   IOField "Default" at 10,10 size 100x30
   TextField "Label_Default" at 10,42 size 67x22; Text 'Default'
   IOField "AboveUpperLimitColor" at 120,10 size 100x30
   TextField "Label_AboveUpperLimitColor" at 120,42 size 194x22; Text 'AboveUpperLimitColor'
   IOField "BackColor" at 230,10 size 100x30
   TextField "Label_BackColor" at 230,42 size 90x22; Text 'BackColor'
   IOField "BackFillStyle" at 340,10 size 100x30
   TextField "Label_BackFillStyle" at 340,42 size 117x22; Text 'BackFillStyle'
   IOField "BelowLowerLimitColor" at 450,10 size 100x30
   TextField "Label_BelowLowerLimitColor" at 450,42 size 196x22; Text 'BelowLowerLimitColor'
   IOField "BorderBackColor" at 560,10 size 100x30
   TextField "Label_BorderBackColor" at 560,42 size 147x22; Text 'BorderBackColor'
   IOField "BorderColor" at 670,10 size 100x30
   TextField "Label_BorderColor" at 670,42 size 107x22; Text 'BorderColor'
   IOField "BorderWidth" at 780,10 size 100x30
   TextField "Label_BorderWidth" at 780,42 size 111x22; Text 'BorderWidth'
   IOField "BottomMargin" at 890,10 size 100x30
   TextField "Label_BottomMargin" at 890,42 size 122x22; Text 'BottomMargin'
   IOField "CornerRadius" at 1000,10 size 100x30
   TextField "Label_CornerRadius" at 1000,42 size 119x22; Text 'CornerRadius'
   IOField "DataFormat_3" at 1110,10 size 100x30
   TextField "Label_DataFormat_3" at 1110,42 size 125x22; Text 'DataFormat_3'
   IOField "EdgeStyle" at 10,66 size 100x30
   TextField "Label_EdgeStyle" at 10,98 size 89x22; Text 'EdgeStyle'
   IOField "EdgeStyle_2" at 120,66 size 100x30
   TextField "Label_EdgeStyle_2" at 120,98 size 111x22; Text 'EdgeStyle_2'
   IOField "EdgeStyle_3" at 230,66 size 100x30
   TextField "Label_EdgeStyle_3" at 230,98 size 111x22; Text 'EdgeStyle_3'
   IOField "EdgeStyle_4" at 340,66 size 100x30
   TextField "Label_EdgeStyle_4" at 340,98 size 111x22; Text 'EdgeStyle_4'
   IOField "FieldLength" at 450,66 size 100x30
   TextField "Label_FieldLength" at 450,98 size 104x22; Text 'FieldLength'
   IOField "FitToLargest" at 560,66 size 92x30
   TextField "Label_FitToLargest" at 560,98 size 112x22; Text 'FitToLargest'
   IOField "Flashing" at 670,66 size 100x30
   TextField "Label_Flashing" at 670,98 size 76x22; Text 'Flashing'
   IOField "ForeColor" at 780,66 size 100x30
   TextField "Label_ForeColor" at 780,98 size 88x22; Text 'ForeColor'
   IOField "FormatPattern" at 890,66 size 100x30; FormatPattern 99.9
   TextField "Label_FormatPattern" at 890,98 size 127x22; Text 'FormatPattern'
   IOField "HorizontalAlignment" at 1000,66 size 100x30
   TextField "Label_HorizontalAlignment" at 1000,98 size 177x22; Text 'HorizontalAlignment'
   IOField "HorizontalAlignment_2" at 1110,66 size 100x30
   TextField "Label_HorizontalAlignment_2" at 1110,98 size 199x22; Text 'HorizontalAlignment_2'
   IOField "LeftMargin" at 10,122 size 100x30
   TextField "Label_LeftMargin" at 10,154 size 97x22; Text 'LeftMargin'
   IOField "Mode" at 120,122 size 100x30
   TextField "Label_Mode" at 120,154 size 49x22; Text 'Mode'
   IOField "Mode_2" at 230,122 size 100x30
   TextField "Label_Mode_2" at 230,154 size 71x22; Text 'Mode_2'
   IOField "RightMargin" at 340,122 size 100x30
   TextField "Label_RightMargin" at 340,154 size 108x22; Text 'RightMargin'
   IOField "ShiftDecimalPoint" at 450,122 size 100x30
   TextField "Label_ShiftDecimalPoint" at 450,154 size 157x22; Text 'ShiftDecimalPoint'
   IOField "ShowLeadingZeros" at 560,122 size 100x30
   TextField "Label_ShowLeadingZeros" at 560,154 size 163x22; Text 'ShowLeadingZeros'
   IOField "TopMargin" at 670,122 size 100x30
   TextField "Label_TopMargin" at 670,154 size 93x22; Text 'TopMargin'
   IOField "Unit" at 780,122 size 100x30; Unit mm
   TextField "Label_Unit" at 780,154 size 40x22; Text 'Unit'
   IOField "UseDesignColorSchema" at 890,122 size 100x30
   TextField "Label_UseDesignColorSchema" at 890,154 size 202x22; Text 'UseDesignColorSchema'
   IOField "VerticalAlignment" at 1000,122 size 100x30
   TextField "Label_VerticalAlignment" at 1000,154 size 156x22; Text 'VerticalAlignment'
   IOField "VerticalAlignment_2" at 1110,122 size 100x30
   TextField "Label_VerticalAlignment_2" at 1110,154 size 178x22; Text 'VerticalAlignment_2'
   Button "Next" at 1238,776 size 40x22; TextOff 'Text'
      on Click: ActivateScreen("P_Button_1", 0)

screen "P_Button_1" 1280x800
   Button "Default" at 10,10 size 100x40; TextOff 'Text'
   TextField "Label_Default" at 10,52 size 67x22; Text 'Default'
   Button "BackColor" at 120,10 size 100x40; TextOff 'Text'
   TextField "Label_BackColor" at 120,52 size 90x22; Text 'BackColor'
   Button "BackFillStyle" at 230,10 size 100x40; TextOff 'Text'
   TextField "Label_BackFillStyle" at 230,52 size 117x22; Text 'BackFillStyle'
   Button "BorderBackColor" at 340,10 size 100x40; TextOff 'Text'
   TextField "Label_BorderBackColor" at 340,52 size 147x22; Text 'BorderBackColor'
   Button "BorderColor" at 450,10 size 100x40; TextOff 'Text'
   TextField "Label_BorderColor" at 450,52 size 107x22; Text 'BorderColor'
   Button "BorderWidth" at 560,10 size 100x40; TextOff 'Text'
   TextField "Label_BorderWidth" at 560,52 size 111x22; Text 'BorderWidth'
   Button "CornerRadius" at 670,10 size 100x40; TextOff 'Text'
   TextField "Label_CornerRadius" at 670,52 size 119x22; Text 'CornerRadius'
   Button "EdgeStyle" at 780,10 size 100x40; TextOff 'Text'
   TextField "Label_EdgeStyle" at 780,52 size 89x22; Text 'EdgeStyle'
   Button "EdgeStyle_2" at 890,10 size 100x40; TextOff 'Text'
   TextField "Label_EdgeStyle_2" at 890,52 size 111x22; Text 'EdgeStyle_2'
   Button "EdgeStyle_3" at 1000,10 size 100x40; TextOff 'Text'
   TextField "Label_EdgeStyle_3" at 1000,52 size 111x22; Text 'EdgeStyle_3'
   Button "EdgeStyle_4" at 1110,10 size 100x40; TextOff 'Text'
   TextField "Label_EdgeStyle_4" at 1110,52 size 111x22; Text 'EdgeStyle_4'
   Button "FirstGradientColor" at 10,76 size 100x40; TextOff 'Text'
   TextField "Label_FirstGradientColor" at 10,118 size 163x22; Text 'FirstGradientColor'
   Button "FirstGradientOffset" at 120,76 size 100x40; TextOff 'Text'
   TextField "Label_FirstGradientOffset" at 120,118 size 171x22; Text 'FirstGradientOffset'
   Button "FitToLargest" at 230,76 size 41x25; TextOff 'Text'
   TextField "Label_FitToLargest" at 230,118 size 112x22; Text 'FitToLargest'
   Button "Flashing" at 340,76 size 100x40; TextOff 'Text'
   TextField "Label_Flashing" at 340,118 size 76x22; Text 'Flashing'
   Button "FocusColor" at 450,76 size 100x40; TextOff 'Text'
   TextField "Label_FocusColor" at 450,118 size 98x22; Text 'FocusColor'
   Button "FocusWidth" at 560,76 size 100x40; TextOff 'Text'
   TextField "Label_FocusWidth" at 560,118 size 102x22; Text 'FocusWidth'
   Button "ForeColor" at 670,76 size 100x40; TextOff 'Text'
   TextField "Label_ForeColor" at 670,118 size 88x22; Text 'ForeColor'
   Button "HorizontalAlignment" at 780,76 size 100x40; TextOff 'Text'
   TextField "Label_HorizontalAlignment" at 780,118 size 177x22; Text 'HorizontalAlignment'
   Button "HorizontalAlignment_2" at 890,76 size 100x40; TextOff 'Text'
   TextField "Label_HorizontalAlignment_2" at 890,118 size 199x22; Text 'HorizontalAlignment_2'
   Button "HorizontalPictureAlignment" at 1000,76 size 100x40; TextOff 'Text'
   TextField "Label_HorizontalPictureAlignment" at 1000,118 size 238x22; Text 'HorizontalPictureAlignment'
   Button "HorizontalPictureAlignment_2" at 1110,76 size 100x40; TextOff 'Text'
   TextField "Label_HorizontalPictureAlignment_2" at 1110,118 size 260x22; Text 'HorizontalPictureAlignment_2'
   Button "MiddleGradientColor" at 10,142 size 100x40; TextOff 'Text'
   TextField "Label_MiddleGradientColor" at 10,184 size 179x22; Text 'MiddleGradientColor'
   Button "Mode_5" at 120,142 size 100x40; TextOff 'Text'
   TextField "Label_Mode_5" at 120,184 size 71x22; Text 'Mode_5'
   Button "Mode_7" at 230,142 size 100x40; TextOff 'Text'
   TextField "Label_Mode_7" at 230,184 size 71x22; Text 'Mode_7'
   Button "PictureAreaBottomMargin" at 340,142 size 100x40; TextOff 'Text'
   TextField "Label_PictureAreaBottomMargin" at 340,184 size 222x22; Text 'PictureAreaBottomMargin'
   Button "PictureAreaLeftMargin" at 450,142 size 100x40; TextOff 'Text'
   TextField "Label_PictureAreaLeftMargin" at 450,184 size 197x22; Text 'PictureAreaLeftMargin'
   Button "PictureAreaRightMargin" at 560,142 size 100x40; TextOff 'Text'
   TextField "Label_PictureAreaRightMargin" at 560,184 size 208x22; Text 'PictureAreaRightMargin'
   Button "PictureAreaTopMargin" at 670,142 size 100x40; TextOff 'Text'
   TextField "Label_PictureAreaTopMargin" at 670,184 size 193x22; Text 'PictureAreaTopMargin'
   Button "SecondGradientColor" at 780,142 size 100x40; TextOff 'Text'
   TextField "Label_SecondGradientColor" at 780,184 size 183x22; Text 'SecondGradientColor'
   Button "SecondGradientOffset" at 890,142 size 100x40; TextOff 'Text'
   TextField "Label_SecondGradientOffset" at 890,184 size 191x22; Text 'SecondGradientOffset'
   Button "TextAreaBottomMargin" at 1000,142 size 100x40; TextOff 'Text'
   TextField "Label_TextAreaBottomMargin" at 1000,184 size 198x22; Text 'TextAreaBottomMargin'
   Button "TextAreaLeftMargin" at 1110,142 size 100x40; TextOff 'Text'
   TextField "Label_TextAreaLeftMargin" at 1110,184 size 173x22; Text 'TextAreaLeftMargin'
   Button "TextAreaRightMargin" at 10,208 size 100x40; TextOff 'Text'
   TextField "Label_TextAreaRightMargin" at 10,250 size 184x22; Text 'TextAreaRightMargin'
   Button "TextAreaTopMargin" at 120,208 size 100x40; TextOff 'Text'
   TextField "Label_TextAreaTopMargin" at 120,250 size 169x22; Text 'TextAreaTopMargin'
   Button "UseDesignColorSchema" at 230,208 size 100x40; TextOff 'Text'
   TextField "Label_UseDesignColorSchema" at 230,250 size 202x22; Text 'UseDesignColorSchema'
   Button "UseFirstGradient" at 340,208 size 100x40; TextOff 'Text'
   TextField "Label_UseFirstGradient" at 340,250 size 149x22; Text 'UseFirstGradient'
   Button "UseSecondGradient" at 450,208 size 100x40; TextOff 'Text'
   TextField "Label_UseSecondGradient" at 450,250 size 169x22; Text 'UseSecondGradient'
   Button "VerticalAlignment" at 560,208 size 100x40; TextOff 'Text'
   TextField "Label_VerticalAlignment" at 560,250 size 156x22; Text 'VerticalAlignment'
   Button "VerticalAlignment_2" at 670,208 size 100x40; TextOff 'Text'
   TextField "Label_VerticalAlignment_2" at 670,250 size 178x22; Text 'VerticalAlignment_2'
   Button "VerticalPictureAlignment" at 780,208 size 100x40; TextOff 'Text'
   TextField "Label_VerticalPictureAlignment" at 780,250 size 217x22; Text 'VerticalPictureAlignment'
   Button "VerticalPictureAlignment_2" at 890,208 size 100x40; TextOff 'Text'
   TextField "Label_VerticalPictureAlignment_2" at 890,250 size 239x22; Text 'VerticalPictureAlignment_2'
   Button "Next" at 1238,776 size 40x22; TextOff 'Text'
      on Click: ActivateScreen("P_SymbolicIOField_1", 0)

screen "P_SymbolicIOField_1" 1280x800
   SymbolicIOField "Default" at 10,10 size 120x30; TextOff '0'; TextOn '1'
   TextField "Label_Default" at 10,42 size 67x22; Text 'Default'
   SymbolicIOField "AboveUpperLimitColor" at 140,10 size 120x30; TextOff '0'; TextOn '1'
   TextField "Label_AboveUpperLimitColor" at 140,42 size 194x22; Text 'AboveUpperLimitColor'
   SymbolicIOField "BackColor" at 270,10 size 120x30; TextOff '0'; TextOn '1'
   TextField "Label_BackColor" at 270,42 size 90x22; Text 'BackColor'
   SymbolicIOField "BackFillStyle" at 400,10 size 120x30; TextOff '0'; TextOn '1'
   TextField "Label_BackFillStyle" at 400,42 size 117x22; Text 'BackFillStyle'
   SymbolicIOField "BelowLowerLimitColor" at 530,10 size 120x30; TextOff '0'; TextOn '1'
   TextField "Label_BelowLowerLimitColor" at 530,42 size 196x22; Text 'BelowLowerLimitColor'
   SymbolicIOField "BorderBackColor" at 660,10 size 120x30; TextOff '0'; TextOn '1'
   TextField "Label_BorderBackColor" at 660,42 size 147x22; Text 'BorderBackColor'
   SymbolicIOField "BorderColor" at 790,10 size 120x30; TextOff '0'; TextOn '1'
   TextField "Label_BorderColor" at 790,42 size 107x22; Text 'BorderColor'
   SymbolicIOField "BorderWidth" at 920,10 size 120x30; TextOff '0'; TextOn '1'
   TextField "Label_BorderWidth" at 920,42 size 111x22; Text 'BorderWidth'
   SymbolicIOField "BottomMargin" at 1050,10 size 120x30; TextOff '0'; TextOn '1'
   TextField "Label_BottomMargin" at 1050,42 size 122x22; Text 'BottomMargin'
   SymbolicIOField "CornerRadius" at 10,66 size 120x30; TextOff '0'; TextOn '1'
   TextField "Label_CornerRadius" at 10,98 size 119x22; Text 'CornerRadius'
   SymbolicIOField "CountVisibleItems" at 140,66 size 120x30; TextOff '0'; TextOn '1'
   TextField "Label_CountVisibleItems" at 140,98 size 159x22; Text 'CountVisibleItems'
   SymbolicIOField "EdgeStyle" at 270,66 size 120x30; TextOff '0'; TextOn '1'
   TextField "Label_EdgeStyle" at 270,98 size 89x22; Text 'EdgeStyle'
   SymbolicIOField "EdgeStyle_2" at 400,66 size 120x30; TextOff '0'; TextOn '1'
   TextField "Label_EdgeStyle_2" at 400,98 size 111x22; Text 'EdgeStyle_2'
   SymbolicIOField "EdgeStyle_3" at 530,66 size 120x30; TextOff '0'; TextOn '1'
   TextField "Label_EdgeStyle_3" at 530,98 size 111x22; Text 'EdgeStyle_3'
   SymbolicIOField "EdgeStyle_4" at 660,66 size 120x30; TextOff '0'; TextOn '1'
   TextField "Label_EdgeStyle_4" at 660,98 size 111x22; Text 'EdgeStyle_4'
   SymbolicIOField "EvenRowBackColor" at 790,66 size 120x30; TextOff '0'; TextOn '1'
   TextField "Label_EvenRowBackColor" at 790,98 size 166x22; Text 'EvenRowBackColor'
   SymbolicIOField "FitToLargest" at 920,66 size 52x30; TextOff '0'; TextOn '1'
   TextField "Label_FitToLargest" at 920,98 size 112x22; Text 'FitToLargest'
   SymbolicIOField "Flashing" at 1050,66 size 120x30; TextOff '0'; TextOn '1'
   TextField "Label_Flashing" at 1050,98 size 76x22; Text 'Flashing'
   SymbolicIOField "FlashingOnLimitViolation" at 10,122 size 120x30; TextOff '0'; TextOn '1'
   TextField "Label_FlashingOnLimitViolation" at 10,154 size 218x22; Text 'FlashingOnLimitViolation'
   SymbolicIOField "ForeColor" at 140,122 size 120x30; TextOff '0'; TextOn '1'
   TextField "Label_ForeColor" at 140,154 size 88x22; Text 'ForeColor'
   SymbolicIOField "HorizontalAlignment" at 270,122 size 120x30; TextOff '0'; TextOn '1'
   TextField "Label_HorizontalAlignment" at 270,154 size 177x22; Text 'HorizontalAlignment'
   SymbolicIOField "HorizontalAlignment_2" at 400,122 size 120x30; TextOff '0'; TextOn '1'
   TextField "Label_HorizontalAlignment_2" at 400,154 size 199x22; Text 'HorizontalAlignment_2'
   SymbolicIOField "LeftMargin" at 530,122 size 120x30; TextOff '0'; TextOn '1'
   TextField "Label_LeftMargin" at 530,154 size 97x22; Text 'LeftMargin'
   SymbolicIOField "Mode" at 660,122 size 120x30; TextOff '0'; TextOn '1'
   TextField "Label_Mode" at 660,154 size 49x22; Text 'Mode'
   SymbolicIOField "Mode_2" at 790,122 size 120x30; TextOff '0'; TextOn '1'
   TextField "Label_Mode_2" at 790,154 size 71x22; Text 'Mode_2'
   SymbolicIOField "RightMargin" at 920,122 size 120x30; TextOff '0'; TextOn '1'
   TextField "Label_RightMargin" at 920,154 size 108x22; Text 'RightMargin'
   SymbolicIOField "SelectBackColor" at 1050,122 size 120x30; TextOff '0'; TextOn '1'
   TextField "Label_SelectBackColor" at 1050,154 size 143x22; Text 'SelectBackColor'
   SymbolicIOField "SelectForeColor" at 10,178 size 120x30; TextOff '0'; TextOn '1'
   TextField "Label_SelectForeColor" at 10,210 size 141x22; Text 'SelectForeColor'
   SymbolicIOField "ShowDropDownButton" at 140,178 size 120x30; TextOff '0'; TextOn '1'
   TextField "Label_ShowDropDownButton" at 140,210 size 191x22; Text 'ShowDropDownButton'
   SymbolicIOField "ShowDropDownList" at 270,178 size 120x30; TextOff '0'; TextOn '1'
   TextField "Label_ShowDropDownList" at 270,210 size 168x22; Text 'ShowDropDownList'
   SymbolicIOField "TopMargin" at 400,178 size 120x30; TextOff '0'; TextOn '1'
   TextField "Label_TopMargin" at 400,210 size 93x22; Text 'TopMargin'
   SymbolicIOField "UseDesignColorSchema" at 530,178 size 120x30; TextOff '0'; TextOn '1'
   TextField "Label_UseDesignColorSchema" at 530,210 size 202x22; Text 'UseDesignColorSchema'
   SymbolicIOField "VerticalAlignment" at 660,178 size 120x30; TextOff '0'; TextOn '1'
   TextField "Label_VerticalAlignment" at 660,210 size 156x22; Text 'VerticalAlignment'
   SymbolicIOField "VerticalAlignment_2" at 790,178 size 120x30; TextOff '0'; TextOn '1'
   TextField "Label_VerticalAlignment_2" at 790,210 size 178x22; Text 'VerticalAlignment_2'
   Button "Next" at 1238,776 size 40x22; TextOff 'Text'
      on Click: ActivateScreen("P_GraphicIOField_1", 0)

screen "P_GraphicIOField_1" 1280x800
   GraphicIOField "Default" at 10,10 size 60x60
   TextField "Label_Default" at 10,72 size 67x22; Text 'Default'
   GraphicIOField "AboveUpperLimitColor" at 80,10 size 60x60
   TextField "Label_AboveUpperLimitColor" at 80,72 size 194x22; Text 'AboveUpperLimitColor'
   GraphicIOField "BackColor" at 150,10 size 60x60
   TextField "Label_BackColor" at 150,72 size 90x22; Text 'BackColor'
   GraphicIOField "BackFillStyle" at 220,10 size 60x60
   TextField "Label_BackFillStyle" at 220,72 size 117x22; Text 'BackFillStyle'
   GraphicIOField "BelowLowerLimitColor" at 290,10 size 60x60
   TextField "Label_BelowLowerLimitColor" at 290,72 size 196x22; Text 'BelowLowerLimitColor'
   GraphicIOField "BorderColor" at 360,10 size 60x60
   TextField "Label_BorderColor" at 360,72 size 107x22; Text 'BorderColor'
   GraphicIOField "BorderWidth" at 430,10 size 60x60
   TextField "Label_BorderWidth" at 430,72 size 111x22; Text 'BorderWidth'
   GraphicIOField "EdgeStyle" at 500,10 size 60x60
   TextField "Label_EdgeStyle" at 500,72 size 89x22; Text 'EdgeStyle'
   GraphicIOField "EdgeStyle_2" at 570,10 size 60x60
   TextField "Label_EdgeStyle_2" at 570,72 size 111x22; Text 'EdgeStyle_2'
   GraphicIOField "EdgeStyle_3" at 640,10 size 60x60
   TextField "Label_EdgeStyle_3" at 640,72 size 111x22; Text 'EdgeStyle_3'
   GraphicIOField "EdgeStyle_4" at 710,10 size 60x60
   TextField "Label_EdgeStyle_4" at 710,72 size 111x22; Text 'EdgeStyle_4'
   GraphicIOField "FitToLargest" at 780,10 size 60x60
   TextField "Label_FitToLargest" at 780,72 size 112x22; Text 'FitToLargest'
   GraphicIOField "Flashing" at 850,10 size 60x60
   TextField "Label_Flashing" at 850,72 size 76x22; Text 'Flashing'
   GraphicIOField "FlashingOnLimitViolation" at 920,10 size 60x60
   TextField "Label_FlashingOnLimitViolation" at 920,72 size 218x22; Text 'FlashingOnLimitViolation'
   GraphicIOField "FocusColor" at 990,10 size 60x60
   TextField "Label_FocusColor" at 990,72 size 98x22; Text 'FocusColor'
   GraphicIOField "FocusWidth" at 1060,10 size 60x60
   TextField "Label_FocusWidth" at 1060,72 size 102x22; Text 'FocusWidth'
   GraphicIOField "Mode" at 1130,10 size 60x60
   TextField "Label_Mode" at 1130,72 size 49x22; Text 'Mode'
   GraphicIOField "Mode_2" at 1200,10 size 60x60
   TextField "Label_Mode_2" at 1200,72 size 71x22; Text 'Mode_2'
   GraphicIOField "ScrollBarOrientation" at 10,96 size 60x60
   TextField "Label_ScrollBarOrientation" at 10,158 size 181x22; Text 'ScrollBarOrientation'
   GraphicIOField "TransparentColor" at 80,96 size 60x60
   TextField "Label_TransparentColor" at 80,158 size 152x22; Text 'TransparentColor'
   GraphicIOField "UseTransparentColor" at 150,96 size 60x60
   TextField "Label_UseTransparentColor" at 150,158 size 183x22; Text 'UseTransparentColor'
   Button "Next" at 1238,776 size 40x22; TextOff 'Text'
      on Click: ActivateScreen("P_DateTimeField_1", 0)

screen "P_DateTimeField_1" 1280x800
   DateTimeField "Default" at 10,10 size 189x26
   TextField "Label_Default" at 10,42 size 67x22; Text 'Default'
   DateTimeField "BackColor" at 180,10 size 189x26
   TextField "Label_BackColor" at 180,42 size 90x22; Text 'BackColor'
   DateTimeField "BackFillStyle" at 350,10 size 189x26
   TextField "Label_BackFillStyle" at 350,42 size 117x22; Text 'BackFillStyle'
   DateTimeField "BorderBackColor" at 520,10 size 189x26
   TextField "Label_BorderBackColor" at 520,42 size 147x22; Text 'BorderBackColor'
   DateTimeField "BorderColor" at 690,10 size 189x26
   TextField "Label_BorderColor" at 690,42 size 107x22; Text 'BorderColor'
   DateTimeField "BorderWidth" at 860,10 size 195x32
   TextField "Label_BorderWidth" at 860,42 size 111x22; Text 'BorderWidth'
   DateTimeField "BottomMargin" at 1030,10 size 189x32
   TextField "Label_BottomMargin" at 1030,42 size 122x22; Text 'BottomMargin'
   DateTimeField "CornerRadius" at 10,66 size 189x26
   TextField "Label_CornerRadius" at 10,98 size 119x22; Text 'CornerRadius'
   DateTimeField "DisplaySystemTime" at 180,66 size 189x26
   TextField "Label_DisplaySystemTime" at 180,98 size 169x22; Text 'DisplaySystemTime'
   DateTimeField "EdgeStyle" at 350,66 size 189x26
   TextField "Label_EdgeStyle" at 350,98 size 89x22; Text 'EdgeStyle'
   DateTimeField "EdgeStyle_2" at 520,66 size 189x26
   TextField "Label_EdgeStyle_2" at 520,98 size 111x22; Text 'EdgeStyle_2'
   DateTimeField "EdgeStyle_3" at 690,66 size 189x26
   TextField "Label_EdgeStyle_3" at 690,98 size 111x22; Text 'EdgeStyle_3'
   DateTimeField "EdgeStyle_4" at 860,66 size 189x26
   TextField "Label_EdgeStyle_4" at 860,98 size 111x22; Text 'EdgeStyle_4'
   DateTimeField "FitToLargest" at 1030,66 size 160x30
   TextField "Label_FitToLargest" at 1030,98 size 112x22; Text 'FitToLargest'
   DateTimeField "Flashing" at 10,122 size 189x26
   TextField "Label_Flashing" at 10,154 size 76x22; Text 'Flashing'
   DateTimeField "ForeColor" at 180,122 size 189x26
   TextField "Label_ForeColor" at 180,154 size 88x22; Text 'ForeColor'
   DateTimeField "HorizontalAlignment" at 350,122 size 189x26
   TextField "Label_HorizontalAlignment" at 350,154 size 177x22; Text 'HorizontalAlignment'
   DateTimeField "HorizontalAlignment_2" at 520,122 size 189x26
   TextField "Label_HorizontalAlignment_2" at 520,154 size 199x22; Text 'HorizontalAlignment_2'
   DateTimeField "LeftMargin" at 690,122 size 195x26
   TextField "Label_LeftMargin" at 690,154 size 97x22; Text 'LeftMargin'
   DateTimeField "LongDateTimeFormat" at 860,122 size 340x26
   TextField "Label_LongDateTimeFormat" at 860,154 size 183x22; Text 'LongDateTimeFormat'
   DateTimeField "Mode_3" at 1030,122 size 189x26
   TextField "Label_Mode_3" at 1030,154 size 71x22; Text 'Mode_3'
   DateTimeField "RightMargin" at 10,178 size 195x26
   TextField "Label_RightMargin" at 10,210 size 108x22; Text 'RightMargin'
   DateTimeField "ShowDate" at 180,178 size 100x26
   TextField "Label_ShowDate" at 180,210 size 89x22; Text 'ShowDate'
   DateTimeField "ShowTime" at 350,178 size 90x26
   TextField "Label_ShowTime" at 350,210 size 90x22; Text 'ShowTime'
   DateTimeField "TopMargin" at 520,178 size 189x32
   TextField "Label_TopMargin" at 520,210 size 93x22; Text 'TopMargin'
   DateTimeField "UseDesignColorSchema" at 690,178 size 234x31
   TextField "Label_UseDesignColorSchema" at 690,210 size 202x22; Text 'UseDesignColorSchema'
   DateTimeField "VerticalAlignment" at 860,178 size 189x26
   TextField "Label_VerticalAlignment" at 860,210 size 156x22; Text 'VerticalAlignment'
   DateTimeField "VerticalAlignment_2" at 1030,178 size 189x26
   TextField "Label_VerticalAlignment_2" at 1030,210 size 178x22; Text 'VerticalAlignment_2'
   Button "Next" at 1238,776 size 40x22; TextOff 'Text'
      on Click: ActivateScreen("P_Bar_1", 0)

screen "P_Bar_1" 1280x800
   Bar "Default" at 10,10 size 40x120
   TextField "Label_Default" at 10,132 size 67x22; Text 'Default'
   Bar "BackColor" at 60,10 size 40x120
   TextField "Label_BackColor" at 60,132 size 90x22; Text 'BackColor'
   Bar "BarBackColor" at 110,10 size 40x120
   TextField "Label_BarBackColor" at 110,132 size 119x22; Text 'BarBackColor'
   Bar "BarEdgeStyle" at 160,10 size 40x120
   TextField "Label_BarEdgeStyle" at 160,132 size 118x22; Text 'BarEdgeStyle'
   Bar "BarEdgeStyle_2" at 210,10 size 40x120
   TextField "Label_BarEdgeStyle_2" at 210,132 size 140x22; Text 'BarEdgeStyle_2'
   Bar "BarOrientation" at 260,10 size 40x120
   TextField "Label_BarOrientation" at 260,132 size 131x22; Text 'BarOrientation'
   Bar "BarOrientation_2" at 310,10 size 40x120
   TextField "Label_BarOrientation_2" at 310,132 size 153x22; Text 'BarOrientation_2'
   Bar "BarOrientation_3" at 360,10 size 40x120
   TextField "Label_BarOrientation_3" at 360,132 size 153x22; Text 'BarOrientation_3'
   Bar "BorderBackColor" at 410,10 size 40x120
   TextField "Label_BorderBackColor" at 410,132 size 147x22; Text 'BorderBackColor'
   Bar "BorderColor" at 460,10 size 40x120
   TextField "Label_BorderColor" at 460,132 size 107x22; Text 'BorderColor'
   Bar "BorderWidth" at 510,10 size 40x120
   TextField "Label_BorderWidth" at 510,132 size 111x22; Text 'BorderWidth'
   Bar "CornerRadius" at 560,10 size 40x120
   TextField "Label_CornerRadius" at 560,132 size 119x22; Text 'CornerRadius'
   Bar "CountSubDivisions" at 610,10 size 40x120
   TextField "Label_CountSubDivisions" at 610,132 size 162x22; Text 'CountSubDivisions'
   Bar "EdgeStyle" at 660,10 size 40x120
   TextField "Label_EdgeStyle" at 660,132 size 89x22; Text 'EdgeStyle'
   Bar "EdgeStyle_2" at 710,10 size 40x120
   TextField "Label_EdgeStyle_2" at 710,132 size 111x22; Text 'EdgeStyle_2'
   Bar "EdgeStyle_3" at 760,10 size 40x120
   TextField "Label_EdgeStyle_3" at 760,132 size 111x22; Text 'EdgeStyle_3'
   Bar "EdgeStyle_4" at 810,10 size 40x120
   TextField "Label_EdgeStyle_4" at 810,132 size 111x22; Text 'EdgeStyle_4'
   Bar "Flashing" at 860,10 size 40x120
   TextField "Label_Flashing" at 860,132 size 76x22; Text 'Flashing'
   Bar "FlashingOnLimitViolation" at 910,10 size 40x120
   TextField "Label_FlashingOnLimitViolation" at 910,132 size 218x22; Text 'FlashingOnLimitViolation'
   Bar "ForeColor" at 960,10 size 40x120
   TextField "Label_ForeColor" at 960,132 size 88x22; Text 'ForeColor'
   Bar "IntegerDigits" at 1010,10 size 40x120
   TextField "Label_IntegerDigits" at 1010,132 size 118x22; Text 'IntegerDigits'
   Bar "LargeTickLabelingStep" at 1060,10 size 40x120
   TextField "Label_LargeTickLabelingStep" at 1060,132 size 198x22; Text 'LargeTickLabelingStep'
   Bar "MaximumValue" at 1110,10 size 40x120; MaximumValue 200
   TextField "Label_MaximumValue" at 1110,132 size 130x22; Text 'MaximumValue'
   Bar "MinimumValue" at 1160,10 size 40x120; MinimumValue -100
   TextField "Label_MinimumValue" at 1160,132 size 126x22; Text 'MinimumValue'
   Bar "Precision" at 1210,10 size 40x120
   TextField "Label_Precision" at 1210,132 size 84x22; Text 'Precision'
   Bar "RangeLower1Color" at 10,156 size 40x120
   TextField "Label_RangeLower1Color" at 10,278 size 165x22; Text 'RangeLower1Color'
   Bar "RangeLower1Enabled" at 60,156 size 40x120
   TextField "Label_RangeLower1Enabled" at 60,278 size 186x22; Text 'RangeLower1Enabled'
   Bar "RangeLower2Color" at 110,156 size 40x120
   TextField "Label_RangeLower2Color" at 110,278 size 165x22; Text 'RangeLower2Color'
   Bar "RangeLower2Enabled" at 160,156 size 40x120
   TextField "Label_RangeLower2Enabled" at 160,278 size 186x22; Text 'RangeLower2Enabled'
   Bar "RangeNormalColor" at 210,156 size 40x120
   TextField "Label_RangeNormalColor" at 210,278 size 163x22; Text 'RangeNormalColor'
   Bar "RangeNormalEnabled" at 260,156 size 40x120
   TextField "Label_RangeNormalEnabled" at 260,278 size 184x22; Text 'RangeNormalEnabled'
   Bar "RangeUpper1Color" at 310,156 size 40x120
   TextField "Label_RangeUpper1Color" at 310,278 size 163x22; Text 'RangeUpper1Color'
   Bar "RangeUpper1Enabled" at 360,156 size 40x120
   TextField "Label_RangeUpper1Enabled" at 360,278 size 184x22; Text 'RangeUpper1Enabled'
   Bar "RangeUpper2Color" at 410,156 size 40x120
   TextField "Label_RangeUpper2Color" at 410,278 size 163x22; Text 'RangeUpper2Color'
   Bar "RangeUpper2Enabled" at 460,156 size 40x120
   TextField "Label_RangeUpper2Enabled" at 460,278 size 184x22; Text 'RangeUpper2Enabled'
   Bar "ScaleColor" at 510,156 size 40x120
   TextField "Label_ScaleColor" at 510,278 size 96x22; Text 'ScaleColor'
   Bar "ScaleGradation" at 560,156 size 40x120
   TextField "Label_ScaleGradation" at 560,278 size 134x22; Text 'ScaleGradation'
   Bar "ScaleLabelingDoubleLined" at 610,156 size 40x120
   TextField "Label_ScaleLabelingDoubleLined" at 610,278 size 227x22; Text 'ScaleLabelingDoubleLined'
   Bar "ScalePosition" at 660,156 size 40x120
   TextField "Label_ScalePosition" at 660,278 size 120x22; Text 'ScalePosition'
   Bar "SegmentColoring" at 710,156 size 40x120
   TextField "Label_SegmentColoring" at 710,278 size 148x22; Text 'SegmentColoring'
   Bar "ShowLimitLines" at 760,156 size 40x120
   TextField "Label_ShowLimitLines" at 760,278 size 138x22; Text 'ShowLimitLines'
   Bar "ShowLimitMarkers" at 810,156 size 40x120
   TextField "Label_ShowLimitMarkers" at 810,278 size 162x22; Text 'ShowLimitMarkers'
   Bar "ShowLimitRanges" at 860,156 size 40x120
   TextField "Label_ShowLimitRanges" at 860,278 size 154x22; Text 'ShowLimitRanges'
   Bar "ShowProcessValue" at 910,156 size 40x120
   TextField "Label_ShowProcessValue" at 910,278 size 163x22; Text 'ShowProcessValue'
   Bar "ShowScale" at 960,156 size 40x120
   TextField "Label_ShowScale" at 960,278 size 96x22; Text 'ShowScale'
   Bar "ShowTickLabels" at 1010,156 size 40x120
   TextField "Label_ShowTickLabels" at 1010,278 size 140x22; Text 'ShowTickLabels'
   Bar "Unit" at 1060,156 size 40x120; Unit mm
   TextField "Label_Unit" at 1060,278 size 40x22; Text 'Unit'
   Bar "UseAutoScaling" at 1110,156 size 40x120
   TextField "Label_UseAutoScaling" at 1110,278 size 136x22; Text 'UseAutoScaling'
   Bar "UseDesignColorSchema" at 1160,156 size 40x120
   TextField "Label_UseDesignColorSchema" at 1160,278 size 202x22; Text 'UseDesignColorSchema'
   Bar "UseExponentialFormat" at 1210,156 size 40x120
   TextField "Label_UseExponentialFormat" at 1210,278 size 194x22; Text 'UseExponentialFormat'
   Button "Next" at 1238,776 size 40x22; TextOff 'Text'
      on Click: ActivateScreen("P_Switch_1", 0)

screen "P_Switch_1" 1280x800
   Switch "Default" at 10,10 size 120x40; CaptionText 'Switch'; TextOff '0'; TextOn '1'
   TextField "Label_Default" at 10,52 size 67x22; Text 'Default'
   Switch "AboveUpperLimitColor" at 140,10 size 120x40; CaptionText 'Switch'; TextOff '0'; TextOn '1'
   TextField "Label_AboveUpperLimitColor" at 140,52 size 194x22; Text 'AboveUpperLimitColor'
   Switch "BackColor" at 270,10 size 120x40; CaptionText 'Switch'; TextOff '0'; TextOn '1'
   TextField "Label_BackColor" at 270,52 size 90x22; Text 'BackColor'
   Switch "BackFillStyle" at 400,10 size 120x40; CaptionText 'Switch'; TextOff '0'; TextOn '1'
   TextField "Label_BackFillStyle" at 400,52 size 117x22; Text 'BackFillStyle'
   Switch "BelowLowerLimitColor" at 530,10 size 120x40; CaptionText 'Switch'; TextOff '0'; TextOn '1'
   TextField "Label_BelowLowerLimitColor" at 530,52 size 196x22; Text 'BelowLowerLimitColor'
   Switch "BorderBackColor" at 660,10 size 120x40; CaptionText 'Switch'; TextOff '0'; TextOn '1'
   TextField "Label_BorderBackColor" at 660,52 size 147x22; Text 'BorderBackColor'
   Switch "BorderColor" at 790,10 size 120x40; CaptionText 'Switch'; TextOff '0'; TextOn '1'
   TextField "Label_BorderColor" at 790,52 size 107x22; Text 'BorderColor'
   Switch "BorderWidth" at 920,10 size 120x40; CaptionText 'Switch'; TextOff '0'; TextOn '1'
   TextField "Label_BorderWidth" at 920,52 size 111x22; Text 'BorderWidth'
   Switch "CaptionColor" at 1050,10 size 120x40; CaptionText 'Switch'; TextOff '0'; TextOn '1'
   TextField "Label_CaptionColor" at 1050,52 size 114x22; Text 'CaptionColor'
   Switch "CornerRadius" at 10,76 size 120x40; CaptionText 'Switch'; TextOff '0'; TextOn '1'
   TextField "Label_CornerRadius" at 10,118 size 119x22; Text 'CornerRadius'
   Switch "EdgeStyle" at 140,76 size 120x40; CaptionText 'Switch'; TextOff '0'; TextOn '1'
   TextField "Label_EdgeStyle" at 140,118 size 89x22; Text 'EdgeStyle'
   Switch "EdgeStyle_2" at 270,76 size 120x40; CaptionText 'Switch'; TextOff '0'; TextOn '1'
   TextField "Label_EdgeStyle_2" at 270,118 size 111x22; Text 'EdgeStyle_2'
   Switch "EdgeStyle_3" at 400,76 size 120x40; CaptionText 'Switch'; TextOff '0'; TextOn '1'
   TextField "Label_EdgeStyle_3" at 400,118 size 111x22; Text 'EdgeStyle_3'
   Switch "EdgeStyle_4" at 530,76 size 120x40; CaptionText 'Switch'; TextOff '0'; TextOn '1'
   TextField "Label_EdgeStyle_4" at 530,118 size 111x22; Text 'EdgeStyle_4'
   Switch "FirstGradientColor" at 660,76 size 120x40; CaptionText 'Switch'; TextOff '0'; TextOn '1'
   TextField "Label_FirstGradientColor" at 660,118 size 163x22; Text 'FirstGradientColor'
   Switch "FirstGradientOffset" at 790,76 size 120x40; CaptionText 'Switch'; TextOff '0'; TextOn '1'
   TextField "Label_FirstGradientOffset" at 790,118 size 171x22; Text 'FirstGradientOffset'
   Switch "FitToLargest" at 920,76 size 120x40; CaptionText 'Switch'; TextOff '0'; TextOn '1'
   TextField "Label_FitToLargest" at 920,118 size 112x22; Text 'FitToLargest'
   Switch "Flashing" at 1050,76 size 120x40; CaptionText 'Switch'; TextOff '0'; TextOn '1'
   TextField "Label_Flashing" at 1050,118 size 76x22; Text 'Flashing'
   Switch "FlashingOnLimitViolation" at 10,142 size 120x40; CaptionText 'Switch'; TextOff '0'; TextOn '1'
   TextField "Label_FlashingOnLimitViolation" at 10,184 size 218x22; Text 'FlashingOnLimitViolation'
   Switch "FocusColor" at 140,142 size 120x40; CaptionText 'Switch'; TextOff '0'; TextOn '1'
   TextField "Label_FocusColor" at 140,184 size 98x22; Text 'FocusColor'
   Switch "FocusWidth" at 270,142 size 120x40; CaptionText 'Switch'; TextOff '0'; TextOn '1'
   TextField "Label_FocusWidth" at 270,184 size 102x22; Text 'FocusWidth'
   Switch "ForeColor" at 400,142 size 120x40; CaptionText 'Switch'; TextOff '0'; TextOn '1'
   TextField "Label_ForeColor" at 400,184 size 88x22; Text 'ForeColor'
   Switch "HorizontalAlignment" at 530,142 size 120x40; CaptionText 'Switch'; TextOff '0'; TextOn '1'
   TextField "Label_HorizontalAlignment" at 530,184 size 177x22; Text 'HorizontalAlignment'
   Switch "HorizontalAlignment_2" at 660,142 size 120x40; CaptionText 'Switch'; TextOff '0'; TextOn '1'
   TextField "Label_HorizontalAlignment_2" at 660,184 size 199x22; Text 'HorizontalAlignment_2'
   Switch "HorizontalPictureAlignment" at 790,142 size 120x40; CaptionText 'Switch'; TextOff '0'; TextOn '1'
   TextField "Label_HorizontalPictureAlignment" at 790,184 size 238x22; Text 'HorizontalPictureAlignment'
   Switch "HorizontalPictureAlignment_2" at 920,142 size 120x40; CaptionText 'Switch'; TextOff '0'; TextOn '1'
   TextField "Label_HorizontalPictureAlignment_2" at 920,184 size 260x22; Text 'HorizontalPictureAlignment_2'
   Switch "InnerBackColorOff" at 1050,142 size 120x40; CaptionText 'Switch'; TextOff '0'; TextOn '1'
   TextField "Label_InnerBackColorOff" at 1050,184 size 163x22; Text 'InnerBackColorOff'
   Switch "InnerBackColorOn" at 10,208 size 120x40; CaptionText 'Switch'; TextOff '0'; TextOn '1'
   TextField "Label_InnerBackColorOn" at 10,250 size 159x22; Text 'InnerBackColorOn'
   Switch "MiddleGradientColor" at 140,208 size 120x40; CaptionText 'Switch'; TextOff '0'; TextOn '1'
   TextField "Label_MiddleGradientColor" at 140,250 size 179x22; Text 'MiddleGradientColor'
   Switch "PictureAreaBottomMargin" at 270,208 size 120x40; CaptionText 'Switch'; TextOff '0'; TextOn '1'
   TextField "Label_PictureAreaBottomMargin" at 270,250 size 222x22; Text 'PictureAreaBottomMargin'
   Switch "PictureAreaLeftMargin" at 400,208 size 120x40; CaptionText 'Switch'; TextOff '0'; TextOn '1'
   TextField "Label_PictureAreaLeftMargin" at 400,250 size 197x22; Text 'PictureAreaLeftMargin'
   Switch "PictureAreaRightMargin" at 530,208 size 120x40; CaptionText 'Switch'; TextOff '0'; TextOn '1'
   TextField "Label_PictureAreaRightMargin" at 530,250 size 208x22; Text 'PictureAreaRightMargin'
   Switch "PictureAreaTopMargin" at 660,208 size 120x40; CaptionText 'Switch'; TextOff '0'; TextOn '1'
   TextField "Label_PictureAreaTopMargin" at 660,250 size 193x22; Text 'PictureAreaTopMargin'
   Switch "SecondGradientColor" at 790,208 size 120x40; CaptionText 'Switch'; TextOff '0'; TextOn '1'
   TextField "Label_SecondGradientColor" at 790,250 size 183x22; Text 'SecondGradientColor'
   Switch "SecondGradientOffset" at 920,208 size 120x40; CaptionText 'Switch'; TextOff '0'; TextOn '1'
   TextField "Label_SecondGradientOffset" at 920,250 size 191x22; Text 'SecondGradientOffset'
   Switch "ShowCaption" at 1050,208 size 120x40; CaptionText 'Switch'; TextOff '0'; TextOn '1'
   TextField "Label_ShowCaption" at 1050,250 size 114x22; Text 'ShowCaption'
   Switch "SwitchOrientation" at 10,274 size 120x40; CaptionText 'Switch'; TextOff '0'; TextOn '1'
   TextField "Label_SwitchOrientation" at 10,316 size 159x22; Text 'SwitchOrientation'
   Switch "SwitchOrientation_2" at 140,274 size 120x40; CaptionText 'Switch'; TextOff '0'; TextOn '1'
   TextField "Label_SwitchOrientation_2" at 140,316 size 181x22; Text 'SwitchOrientation_2'
   Switch "SwitchOrientation_3" at 270,274 size 120x40; CaptionText 'Switch'; TextOff '0'; TextOn '1'
   TextField "Label_SwitchOrientation_3" at 270,316 size 181x22; Text 'SwitchOrientation_3'
   Switch "TextAreaBottomMargin" at 400,274 size 120x40; CaptionText 'Switch'; TextOff '0'; TextOn '1'
   TextField "Label_TextAreaBottomMargin" at 400,316 size 198x22; Text 'TextAreaBottomMargin'
   Switch "TextAreaLeftMargin" at 530,274 size 120x40; CaptionText 'Switch'; TextOff '0'; TextOn '1'
   TextField "Label_TextAreaLeftMargin" at 530,316 size 173x22; Text 'TextAreaLeftMargin'
   Switch "TextAreaRightMargin" at 660,274 size 120x40; CaptionText 'Switch'; TextOff '0'; TextOn '1'
   TextField "Label_TextAreaRightMargin" at 660,316 size 184x22; Text 'TextAreaRightMargin'
   Switch "TextAreaTopMargin" at 790,274 size 120x40; CaptionText 'Switch'; TextOff '0'; TextOn '1'
   TextField "Label_TextAreaTopMargin" at 790,316 size 169x22; Text 'TextAreaTopMargin'
   Switch "UseDesignColorSchema" at 920,274 size 120x40; CaptionText 'Switch'; TextOff '0'; TextOn '1'
   TextField "Label_UseDesignColorSchema" at 920,316 size 202x22; Text 'UseDesignColorSchema'
   Switch "UseFirstGradient" at 1050,274 size 120x40; CaptionText 'Switch'; TextOff '0'; TextOn '1'
   TextField "Label_UseFirstGradient" at 1050,316 size 149x22; Text 'UseFirstGradient'
   Switch "UseSecondGradient" at 10,340 size 120x40; CaptionText 'Switch'; TextOff '0'; TextOn '1'
   TextField "Label_UseSecondGradient" at 10,382 size 169x22; Text 'UseSecondGradient'
   Switch "VerticalAlignment" at 140,340 size 120x40; CaptionText 'Switch'; TextOff '0'; TextOn '1'
   TextField "Label_VerticalAlignment" at 140,382 size 156x22; Text 'VerticalAlignment'
   Switch "VerticalAlignment_2" at 270,340 size 120x40; CaptionText 'Switch'; TextOff '0'; TextOn '1'
   TextField "Label_VerticalAlignment_2" at 270,382 size 178x22; Text 'VerticalAlignment_2'
   Switch "VerticalPictureAlignment" at 400,340 size 120x40; CaptionText 'Switch'; TextOff '0'; TextOn '1'
   TextField "Label_VerticalPictureAlignment" at 400,382 size 217x22; Text 'VerticalPictureAlignment'
   Switch "VerticalPictureAlignment_2" at 530,340 size 120x40; CaptionText 'Switch'; TextOff '0'; TextOn '1'
   TextField "Label_VerticalPictureAlignment_2" at 530,382 size 239x22; Text 'VerticalPictureAlignment_2'
   Button "Next" at 1238,776 size 40x22; TextOff 'Text'
      on Click: ActivateScreen("P_SymbolLibrary_1", 0)

screen "P_SymbolLibrary_1" 1280x800
   SymbolLibrary "Default" at 10,10 size 60x60
   TextField "Label_Default" at 10,72 size 67x22; Text 'Default'
   SymbolLibrary "AboveUpperLimitColor" at 80,10 size 60x60
   TextField "Label_AboveUpperLimitColor" at 80,72 size 194x22; Text 'AboveUpperLimitColor'
   SymbolLibrary "BackColor" at 150,10 size 60x60
   TextField "Label_BackColor" at 150,72 size 90x22; Text 'BackColor'
   SymbolLibrary "BackFillStyle" at 220,10 size 60x60
   TextField "Label_BackFillStyle" at 220,72 size 117x22; Text 'BackFillStyle'
   SymbolLibrary "BelowLowerLimitColor" at 290,10 size 60x60
   TextField "Label_BelowLowerLimitColor" at 290,72 size 196x22; Text 'BelowLowerLimitColor'
   SymbolLibrary "BlinkColor" at 360,10 size 60x60
   TextField "Label_BlinkColor" at 360,72 size 93x22; Text 'BlinkColor'
   SymbolLibrary "FillColorMode" at 430,10 size 60x60
   TextField "Label_FillColorMode" at 430,72 size 122x22; Text 'FillColorMode'
   SymbolLibrary "FillColorMode_2" at 500,10 size 60x60
   TextField "Label_FillColorMode_2" at 500,72 size 144x22; Text 'FillColorMode_2'
   SymbolLibrary "FixedAspectRatio" at 570,10 size 60x60
   TextField "Label_FixedAspectRatio" at 570,72 size 152x22; Text 'FixedAspectRatio'
   SymbolLibrary "Flashing" at 640,10 size 60x60
   TextField "Label_Flashing" at 640,72 size 76x22; Text 'Flashing'
   SymbolLibrary "FlashingOnLimitViolation" at 710,10 size 60x60
   TextField "Label_FlashingOnLimitViolation" at 710,72 size 218x22; Text 'FlashingOnLimitViolation'
   SymbolLibrary "Flip" at 780,10 size 60x60
   TextField "Label_Flip" at 780,72 size 37x22; Text 'Flip'
   SymbolLibrary "Flip_2" at 850,10 size 60x60
   TextField "Label_Flip_2" at 850,72 size 59x22; Text 'Flip_2'
   SymbolLibrary "Flip_3" at 920,10 size 60x60
   TextField "Label_Flip_3" at 920,72 size 59x22; Text 'Flip_3'
   SymbolLibrary "ForeColor" at 990,10 size 60x60
   TextField "Label_ForeColor" at 990,72 size 88x22; Text 'ForeColor'
   SymbolLibrary "Rotation" at 1060,10 size 60x60
   TextField "Label_Rotation" at 1060,72 size 77x22; Text 'Rotation'
   SymbolLibrary "Rotation_2" at 1130,10 size 60x60
   TextField "Label_Rotation_2" at 1130,72 size 99x22; Text 'Rotation_2'
   SymbolLibrary "Rotation_3" at 1200,10 size 60x60
   TextField "Label_Rotation_3" at 1200,72 size 99x22; Text 'Rotation_3'
   Button "Next" at 1238,776 size 40x22; TextOff 'Text'
      on Click: ActivateScreen("P_Slider_1", 0)

screen "P_Slider_1" 1280x800
   Slider "Default" at 10,10 size 60x160; Caption 'SIMATIC'
   TextField "Label_Default" at 10,172 size 67x22; Text 'Default'
   Slider "BackColor" at 80,10 size 60x160; Caption 'SIMATIC'
   TextField "Label_BackColor" at 80,172 size 90x22; Text 'BackColor'
   Slider "BackFillStyle" at 150,10 size 60x160; Caption 'SIMATIC'
   TextField "Label_BackFillStyle" at 150,172 size 117x22; Text 'BackFillStyle'
   Slider "BarBackColor" at 220,10 size 60x160; Caption 'SIMATIC'
   TextField "Label_BarBackColor" at 220,172 size 119x22; Text 'BarBackColor'
   Slider "BarColor" at 290,10 size 60x160; Caption 'SIMATIC'
   TextField "Label_BarColor" at 290,172 size 79x22; Text 'BarColor'
   Slider "BarOrientation" at 360,10 size 60x160; Caption 'SIMATIC'
   TextField "Label_BarOrientation" at 360,172 size 131x22; Text 'BarOrientation'
   Slider "BarOrientation_2" at 430,10 size 60x160; Caption 'SIMATIC'
   TextField "Label_BarOrientation_2" at 430,172 size 153x22; Text 'BarOrientation_2'
   Slider "BarOrientation_3" at 500,10 size 60x160; Caption 'SIMATIC'
   TextField "Label_BarOrientation_3" at 500,172 size 153x22; Text 'BarOrientation_3'
   Slider "BorderBackColor" at 570,10 size 60x160; Caption 'SIMATIC'
   TextField "Label_BorderBackColor" at 570,172 size 147x22; Text 'BorderBackColor'
   Slider "BorderBrightColor3D" at 640,10 size 60x160; Caption 'SIMATIC'
   TextField "Label_BorderBrightColor3D" at 640,172 size 182x22; Text 'BorderBrightColor3D'
   Slider "BorderColor" at 710,10 size 60x160; Caption 'SIMATIC'
   TextField "Label_BorderColor" at 710,172 size 107x22; Text 'BorderColor'
   Slider "BorderInnerStyle3D" at 780,10 size 60x160; Caption 'SIMATIC'
   TextField "Label_BorderInnerStyle3D" at 780,172 size 175x22; Text 'BorderInnerStyle3D'
   Slider "BorderInnerStyle3D_2" at 850,10 size 60x160; Caption 'SIMATIC'
   TextField "Label_BorderInnerStyle3D_2" at 850,172 size 197x22; Text 'BorderInnerStyle3D_2'
   Slider "BorderInnerWidth3D" at 920,10 size 60x160; Caption 'SIMATIC'
   TextField "Label_BorderInnerWidth3D" at 920,172 size 180x22; Text 'BorderInnerWidth3D'
   Slider "BorderOuterStyle3D" at 990,10 size 60x160; Caption 'SIMATIC'
   TextField "Label_BorderOuterStyle3D" at 990,172 size 177x22; Text 'BorderOuterStyle3D'
   Slider "BorderOuterStyle3D_2" at 1060,10 size 60x160; Caption 'SIMATIC'
   TextField "Label_BorderOuterStyle3D_2" at 1060,172 size 199x22; Text 'BorderOuterStyle3D_2'
   Slider "BorderOuterWidth3D" at 1130,10 size 60x160; Caption 'SIMATIC'
   TextField "Label_BorderOuterWidth3D" at 1130,172 size 182x22; Text 'BorderOuterWidth3D'
   Slider "BorderShadeColor3D" at 1200,10 size 60x160; Caption 'SIMATIC'
   TextField "Label_BorderShadeColor3D" at 1200,172 size 181x22; Text 'BorderShadeColor3D'
   Slider "BorderWidth" at 10,196 size 60x160; Caption 'SIMATIC'
   TextField "Label_BorderWidth" at 10,358 size 111x22; Text 'BorderWidth'
   Slider "CornerRadius" at 80,196 size 60x160; Caption 'SIMATIC'
   TextField "Label_CornerRadius" at 80,358 size 119x22; Text 'CornerRadius'
   Slider "EdgeStyle" at 150,196 size 60x160; Caption 'SIMATIC'
   TextField "Label_EdgeStyle" at 150,358 size 89x22; Text 'EdgeStyle'
   Slider "EdgeStyle_2" at 220,196 size 60x160; Caption 'SIMATIC'
   TextField "Label_EdgeStyle_2" at 220,358 size 111x22; Text 'EdgeStyle_2'
   Slider "EdgeStyle_3" at 290,196 size 60x160; Caption 'SIMATIC'
   TextField "Label_EdgeStyle_3" at 290,358 size 111x22; Text 'EdgeStyle_3'
   Slider "EdgeStyle_4" at 360,196 size 60x160; Caption 'SIMATIC'
   TextField "Label_EdgeStyle_4" at 360,358 size 111x22; Text 'EdgeStyle_4'
   Slider "Flashing" at 430,196 size 60x160; Caption 'SIMATIC'
   TextField "Label_Flashing" at 430,358 size 76x22; Text 'Flashing'
   Slider "FocusColor" at 500,196 size 60x160; Caption 'SIMATIC'
   TextField "Label_FocusColor" at 500,358 size 98x22; Text 'FocusColor'
   Slider "FocusWidth" at 570,196 size 60x160; Caption 'SIMATIC'
   TextField "Label_FocusWidth" at 570,358 size 102x22; Text 'FocusWidth'
   Slider "ForeColor" at 640,196 size 60x160; Caption 'SIMATIC'
   TextField "Label_ForeColor" at 640,358 size 88x22; Text 'ForeColor'
   Slider "LabelColor" at 710,196 size 60x160; Caption 'SIMATIC'
   TextField "Label_LabelColor" at 710,358 size 96x22; Text 'LabelColor'
   Slider "MaximumValue" at 780,196 size 60x160; Caption 'SIMATIC'
   TextField "Label_MaximumValue" at 780,358 size 130x22; Text 'MaximumValue'
   Slider "MinimumValue" at 850,196 size 60x160; Caption 'SIMATIC'
   TextField "Label_MinimumValue" at 850,358 size 126x22; Text 'MinimumValue'
   Slider "RangeLower1Color" at 920,196 size 60x160; Caption 'SIMATIC'
   TextField "Label_RangeLower1Color" at 920,358 size 165x22; Text 'RangeLower1Color'
   Slider "RangeLower1Enabled" at 990,196 size 60x160; Caption 'SIMATIC'
   TextField "Label_RangeLower1Enabled" at 990,358 size 186x22; Text 'RangeLower1Enabled'
   Slider "RangeLower2Color" at 1060,196 size 60x160; Caption 'SIMATIC'
   TextField "Label_RangeLower2Color" at 1060,358 size 165x22; Text 'RangeLower2Color'
   Slider "RangeLower2Enabled" at 1130,196 size 60x160; Caption 'SIMATIC'
   TextField "Label_RangeLower2Enabled" at 1130,358 size 186x22; Text 'RangeLower2Enabled'
   Slider "RangeNormalColor" at 1200,196 size 60x160; Caption 'SIMATIC'
   TextField "Label_RangeNormalColor" at 1200,358 size 163x22; Text 'RangeNormalColor'
   Slider "RangeNormalEnabled" at 10,382 size 60x160; Caption 'SIMATIC'
   TextField "Label_RangeNormalEnabled" at 10,544 size 184x22; Text 'RangeNormalEnabled'
   Slider "RangeUpper1Color" at 80,382 size 60x160; Caption 'SIMATIC'
   TextField "Label_RangeUpper1Color" at 80,544 size 163x22; Text 'RangeUpper1Color'
   Slider "RangeUpper1Enabled" at 150,382 size 60x160; Caption 'SIMATIC'
   TextField "Label_RangeUpper1Enabled" at 150,544 size 184x22; Text 'RangeUpper1Enabled'
   Slider "RangeUpper2Color" at 220,382 size 60x160; Caption 'SIMATIC'
   TextField "Label_RangeUpper2Color" at 220,544 size 163x22; Text 'RangeUpper2Color'
   Slider "RangeUpper2Enabled" at 290,382 size 60x160; Caption 'SIMATIC'
   TextField "Label_RangeUpper2Enabled" at 290,544 size 184x22; Text 'RangeUpper2Enabled'
   Slider "ScalePosition" at 360,382 size 60x160; Caption 'SIMATIC'
   TextField "Label_ScalePosition" at 360,544 size 120x22; Text 'ScalePosition'
   Slider "ShowBar" at 430,382 size 60x160; Caption 'SIMATIC'
   TextField "Label_ShowBar" at 430,544 size 79x22; Text 'ShowBar'
   Slider "ShowLimitLines" at 500,382 size 60x160; Caption 'SIMATIC'
   TextField "Label_ShowLimitLines" at 500,544 size 138x22; Text 'ShowLimitLines'
   Slider "ShowLimitMarkers" at 570,382 size 60x160; Caption 'SIMATIC'
   TextField "Label_ShowLimitMarkers" at 570,544 size 162x22; Text 'ShowLimitMarkers'
   Slider "ShowLimitRanges" at 640,382 size 60x160; Caption 'SIMATIC'
   TextField "Label_ShowLimitRanges" at 640,544 size 154x22; Text 'ShowLimitRanges'
   Slider "ShowPosition" at 710,382 size 60x160; Caption 'SIMATIC'
   TextField "Label_ShowPosition" at 710,544 size 119x22; Text 'ShowPosition'
   Slider "ShowScale" at 780,382 size 60x160; Caption 'SIMATIC'
   TextField "Label_ShowScale" at 780,544 size 96x22; Text 'ShowScale'
   Slider "ShowThumb" at 850,382 size 60x160; Caption 'SIMATIC'
   TextField "Label_ShowThumb" at 850,544 size 104x22; Text 'ShowThumb'
   Slider "ShowTickLabels" at 920,382 size 60x160; Caption 'SIMATIC'
   TextField "Label_ShowTickLabels" at 920,544 size 140x22; Text 'ShowTickLabels'
   Slider "ShowTicks" at 990,382 size 60x160; Caption 'SIMATIC'
   TextField "Label_ShowTicks" at 990,544 size 94x22; Text 'ShowTicks'
   Slider "ThumbBackColor" at 1060,382 size 60x160; Caption 'SIMATIC'
   TextField "Label_ThumbBackColor" at 1060,544 size 144x22; Text 'ThumbBackColor'
   Slider "UseDesignColorSchema" at 1130,382 size 60x160; Caption 'SIMATIC'
   TextField "Label_UseDesignColorSchema" at 1130,544 size 202x22; Text 'UseDesignColorSchema'
   Button "Next" at 1238,776 size 40x22; TextOff 'Text'
      on Click: ActivateScreen("P_Gauge_1", 0)

screen "P_Gauge_1" 1280x800
   Gauge "Default" at 10,10 size 150x150; CaptionText 'SIMATIC'
   TextField "Label_Default" at 10,162 size 67x22; Text 'Default'
   Gauge "AngleMax" at 170,10 size 150x150; CaptionText 'SIMATIC'
   TextField "Label_AngleMax" at 170,162 size 86x22; Text 'AngleMax'
   Gauge "AngleMin" at 330,10 size 150x150; CaptionText 'SIMATIC'
   TextField "Label_AngleMin" at 330,162 size 82x22; Text 'AngleMin'
   Gauge "BackColor" at 490,10 size 150x150; CaptionText 'SIMATIC'
   TextField "Label_BackColor" at 490,162 size 90x22; Text 'BackColor'
   Gauge "BackFillStyle" at 650,10 size 150x150; CaptionText 'SIMATIC'
   TextField "Label_BackFillStyle" at 650,162 size 117x22; Text 'BackFillStyle'
   Gauge "BorderBackColor" at 810,10 size 150x150; CaptionText 'SIMATIC'
   TextField "Label_BorderBackColor" at 810,162 size 147x22; Text 'BorderBackColor'
   Gauge "BorderColor" at 970,10 size 150x150; CaptionText 'SIMATIC'
   TextField "Label_BorderColor" at 970,162 size 107x22; Text 'BorderColor'
   Gauge "BorderWidth" at 10,186 size 150x150; CaptionText 'SIMATIC'
   TextField "Label_BorderWidth" at 10,338 size 111x22; Text 'BorderWidth'
   Gauge "CaptionColor" at 170,186 size 150x150; CaptionText 'SIMATIC'
   TextField "Label_CaptionColor" at 170,338 size 114x22; Text 'CaptionColor'
   Gauge "CaptionTop" at 330,186 size 150x150; CaptionText 'SIMATIC'
   TextField "Label_CaptionTop" at 330,338 size 99x22; Text 'CaptionTop'
   Gauge "CenterColor" at 490,186 size 150x150; CaptionText 'SIMATIC'
   TextField "Label_CenterColor" at 490,338 size 106x22; Text 'CenterColor'
   Gauge "CenterSize" at 650,186 size 150x150; CaptionText 'SIMATIC'
   TextField "Label_CenterSize" at 650,338 size 97x22; Text 'CenterSize'
   Gauge "CornerRadius" at 810,186 size 150x150; CaptionText 'SIMATIC'
   TextField "Label_CornerRadius" at 810,338 size 119x22; Text 'CornerRadius'
   Gauge "DialColor" at 970,186 size 150x150; CaptionText 'SIMATIC'
   TextField "Label_DialColor" at 970,338 size 84x22; Text 'DialColor'
   Gauge "DialFillStyle" at 10,362 size 150x150; CaptionText 'SIMATIC'
   TextField "Label_DialFillStyle" at 10,514 size 111x22; Text 'DialFillStyle'
   Gauge "DialSize" at 170,362 size 150x150; CaptionText 'SIMATIC'
   TextField "Label_DialSize" at 170,514 size 75x22; Text 'DialSize'
   Gauge "EdgeStyle" at 330,362 size 150x150; CaptionText 'SIMATIC'
   TextField "Label_EdgeStyle" at 330,514 size 89x22; Text 'EdgeStyle'
   Gauge "EdgeStyle_2" at 490,362 size 150x150; CaptionText 'SIMATIC'
   TextField "Label_EdgeStyle_2" at 490,514 size 111x22; Text 'EdgeStyle_2'
   Gauge "EdgeStyle_3" at 650,362 size 150x150; CaptionText 'SIMATIC'
   TextField "Label_EdgeStyle_3" at 650,514 size 111x22; Text 'EdgeStyle_3'
   Gauge "EdgeStyle_4" at 810,362 size 150x150; CaptionText 'SIMATIC'
   TextField "Label_EdgeStyle_4" at 810,514 size 111x22; Text 'EdgeStyle_4'
   Gauge "Gradation" at 970,362 size 150x150; CaptionText 'SIMATIC'
   TextField "Label_Gradation" at 970,514 size 88x22; Text 'Gradation'
   Gauge "InnerDialColor" at 10,538 size 150x150; CaptionText 'SIMATIC'
   TextField "Label_InnerDialColor" at 10,690 size 130x22; Text 'InnerDialColor'
   Gauge "InnerDialInnerDistance" at 170,538 size 150x150; CaptionText 'SIMATIC'
   TextField "Label_InnerDialInnerDistance" at 170,690 size 204x22; Text 'InnerDialInnerDistance'
   Gauge "InnerDialOuterDistance" at 330,538 size 150x150; CaptionText 'SIMATIC'
   TextField "Label_InnerDialOuterDistance" at 330,690 size 206x22; Text 'InnerDialOuterDistance'
   Gauge "LockSquaredExtent" at 490,538 size 150x150; CaptionText 'SIMATIC'
   TextField "Label_LockSquaredExtent" at 490,690 size 167x22; Text 'LockSquaredExtent'
   Gauge "MaximumValue" at 650,538 size 150x150; CaptionText 'SIMATIC'
   TextField "Label_MaximumValue" at 650,690 size 130x22; Text 'MaximumValue'
   Gauge "MinimumValue" at 810,538 size 150x150; CaptionText 'SIMATIC'
   TextField "Label_MinimumValue" at 810,690 size 126x22; Text 'MinimumValue'
   Gauge "NeedleHeight" at 970,538 size 150x150; CaptionText 'SIMATIC'
   TextField "Label_NeedleHeight" at 970,690 size 119x22; Text 'NeedleHeight'
   Button "Next" at 1238,776 size 40x22; TextOff 'Text'
      on Click: ActivateScreen("P_Gauge_2", 0)

screen "P_Gauge_2" 1280x800
   Gauge "PointerColor" at 10,10 size 150x150; CaptionText 'SIMATIC'
   TextField "Label_PointerColor" at 10,162 size 112x22; Text 'PointerColor'
   Gauge "RangeLower1Color" at 170,10 size 150x150; CaptionText 'SIMATIC'
   TextField "Label_RangeLower1Color" at 170,162 size 165x22; Text 'RangeLower1Color'
   Gauge "RangeLower1Enabled" at 330,10 size 150x150; CaptionText 'SIMATIC'
   TextField "Label_RangeLower1Enabled" at 330,162 size 186x22; Text 'RangeLower1Enabled'
   Gauge "RangeLower2Color" at 490,10 size 150x150; CaptionText 'SIMATIC'
   TextField "Label_RangeLower2Color" at 490,162 size 165x22; Text 'RangeLower2Color'
   Gauge "RangeLower2Enabled" at 650,10 size 150x150; CaptionText 'SIMATIC'
   TextField "Label_RangeLower2Enabled" at 650,162 size 186x22; Text 'RangeLower2Enabled'
   Gauge "RangeNormalColor" at 810,10 size 150x150; CaptionText 'SIMATIC'
   TextField "Label_RangeNormalColor" at 810,162 size 163x22; Text 'RangeNormalColor'
   Gauge "RangeNormalEnabled" at 970,10 size 150x150; CaptionText 'SIMATIC'
   TextField "Label_RangeNormalEnabled" at 970,162 size 184x22; Text 'RangeNormalEnabled'
   Gauge "RangeUpper1Color" at 10,186 size 150x150; CaptionText 'SIMATIC'
   TextField "Label_RangeUpper1Color" at 10,338 size 163x22; Text 'RangeUpper1Color'
   Gauge "RangeUpper1Enabled" at 170,186 size 150x150; CaptionText 'SIMATIC'
   TextField "Label_RangeUpper1Enabled" at 170,338 size 184x22; Text 'RangeUpper1Enabled'
   Gauge "RangeUpper1Start" at 330,186 size 150x150; CaptionText 'SIMATIC'
   TextField "Label_RangeUpper1Start" at 330,338 size 161x22; Text 'RangeUpper1Start'
   Gauge "RangeUpper2Color" at 490,186 size 150x150; CaptionText 'SIMATIC'
   TextField "Label_RangeUpper2Color" at 490,338 size 163x22; Text 'RangeUpper2Color'
   Gauge "RangeUpper2Enabled" at 650,186 size 150x150; CaptionText 'SIMATIC'
   TextField "Label_RangeUpper2Enabled" at 650,338 size 184x22; Text 'RangeUpper2Enabled'
   Gauge "RangeUpper2Start" at 810,186 size 150x150; CaptionText 'SIMATIC'
   TextField "Label_RangeUpper2Start" at 810,338 size 161x22; Text 'RangeUpper2Start'
   Gauge "ScaleLabelColor" at 970,186 size 150x150; CaptionText 'SIMATIC'
   TextField "Label_ScaleLabelColor" at 970,338 size 142x22; Text 'ScaleLabelColor'
   Gauge "ScaleTickColor" at 10,362 size 150x150; CaptionText 'SIMATIC'
   TextField "Label_ScaleTickColor" at 10,514 size 131x22; Text 'ScaleTickColor'
   Gauge "ScaleTickLabelPosition" at 170,362 size 150x150; CaptionText 'SIMATIC'
   TextField "Label_ScaleTickLabelPosition" at 170,514 size 201x22; Text 'ScaleTickLabelPosition'
   Gauge "ScaleTickLength" at 330,362 size 150x150; CaptionText 'SIMATIC'
   TextField "Label_ScaleTickLength" at 330,514 size 143x22; Text 'ScaleTickLength'
   Gauge "ScaleTickPosition" at 490,362 size 150x150; CaptionText 'SIMATIC'
   TextField "Label_ScaleTickPosition" at 490,514 size 155x22; Text 'ScaleTickPosition'
   Gauge "ShowDecimalPoint" at 650,362 size 150x150; CaptionText 'SIMATIC'
   TextField "Label_ShowDecimalPoint" at 650,514 size 161x22; Text 'ShowDecimalPoint'
   Gauge "ShowInnerDial" at 810,362 size 150x150; CaptionText 'SIMATIC'
   TextField "Label_ShowInnerDial" at 810,514 size 130x22; Text 'ShowInnerDial'
   Gauge "ShowLimitRanges" at 970,362 size 150x150; CaptionText 'SIMATIC'
   TextField "Label_ShowLimitRanges" at 970,514 size 154x22; Text 'ShowLimitRanges'
   Gauge "ShowPeakValuePointer" at 10,538 size 150x150; CaptionText 'SIMATIC'
   TextField "Label_ShowPeakValuePointer" at 10,690 size 200x22; Text 'ShowPeakValuePointer'
   Gauge "UnitColor" at 170,538 size 150x150; CaptionText 'SIMATIC'
   TextField "Label_UnitColor" at 170,690 size 85x22; Text 'UnitColor'
   Gauge "UnitTop" at 330,538 size 150x150; CaptionText 'SIMATIC'
   TextField "Label_UnitTop" at 330,690 size 70x22; Text 'UnitTop'
   Gauge "UseDesignColorSchema" at 490,538 size 150x150; CaptionText 'SIMATIC'
   TextField "Label_UseDesignColorSchema" at 490,690 size 202x22; Text 'UseDesignColorSchema'
   Button "Next" at 1238,776 size 40x22; TextOff 'Text'
      on Click: ActivateScreen("P_Clock_1", 0)

screen "P_Clock_1" 1280x800
   Clock "Default" at 10,10 size 150x150
   TextField "Label_Default" at 10,162 size 67x22; Text 'Default'
   Clock "Analog" at 170,10 size 150x150
   TextField "Label_Analog" at 170,162 size 62x22; Text 'Analog'
   Clock "BackFillStyle" at 330,10 size 150x150
   TextField "Label_BackFillStyle" at 330,162 size 117x22; Text 'BackFillStyle'
   Clock "BorderBackColor" at 490,10 size 150x150
   TextField "Label_BorderBackColor" at 490,162 size 147x22; Text 'BorderBackColor'
   Clock "BorderColor" at 650,10 size 150x150
   TextField "Label_BorderColor" at 650,162 size 107x22; Text 'BorderColor'
   Clock "BorderWidth" at 810,10 size 150x150
   TextField "Label_BorderWidth" at 810,162 size 111x22; Text 'BorderWidth'
   Clock "CornerRadius" at 970,10 size 150x150
   TextField "Label_CornerRadius" at 970,162 size 119x22; Text 'CornerRadius'
   Clock "DialColor" at 10,186 size 150x150
   TextField "Label_DialColor" at 10,338 size 84x22; Text 'DialColor'
   Clock "EdgeStyle" at 170,186 size 150x150
   TextField "Label_EdgeStyle" at 170,338 size 89x22; Text 'EdgeStyle'
   Clock "EdgeStyle_2" at 330,186 size 150x150
   TextField "Label_EdgeStyle_2" at 330,338 size 111x22; Text 'EdgeStyle_2'
   Clock "EdgeStyle_3" at 490,186 size 150x150
   TextField "Label_EdgeStyle_3" at 490,338 size 111x22; Text 'EdgeStyle_3'
   Clock "EdgeStyle_4" at 650,186 size 150x150
   TextField "Label_EdgeStyle_4" at 650,338 size 111x22; Text 'EdgeStyle_4'
   Clock "Flashing" at 810,186 size 150x150
   TextField "Label_Flashing" at 810,338 size 76x22; Text 'Flashing'
   Clock "HourNeedleHeight" at 970,186 size 150x150
   TextField "Label_HourNeedleHeight" at 970,338 size 159x22; Text 'HourNeedleHeight'
   Clock "HourNeedleWidth" at 10,362 size 150x150
   TextField "Label_HourNeedleWidth" at 10,514 size 153x22; Text 'HourNeedleWidth'
   Clock "LockSquaredExtent" at 170,362 size 150x150
   TextField "Label_LockSquaredExtent" at 170,514 size 167x22; Text 'LockSquaredExtent'
   Clock "MinuteNeedleHeight" at 330,362 size 150x150
   TextField "Label_MinuteNeedleHeight" at 330,514 size 176x22; Text 'MinuteNeedleHeight'
   Clock "MinuteNeedleWidth" at 490,362 size 150x150
   TextField "Label_MinuteNeedleWidth" at 490,514 size 170x22; Text 'MinuteNeedleWidth'
   Clock "NeedleBorderColor" at 650,362 size 150x150
   TextField "Label_NeedleBorderColor" at 650,514 size 166x22; Text 'NeedleBorderColor'
   Clock "NeedleColor" at 810,362 size 150x150
   TextField "Label_NeedleColor" at 810,514 size 109x22; Text 'NeedleColor'
   Clock "NeedleFillStyle" at 970,362 size 150x150
   TextField "Label_NeedleFillStyle" at 970,514 size 136x22; Text 'NeedleFillStyle'
   Clock "NumberStyle" at 10,538 size 150x150
   TextField "Label_NumberStyle" at 10,690 size 114x22; Text 'NumberStyle'
   Clock "NumberStyle_2" at 170,538 size 150x150
   TextField "Label_NumberStyle_2" at 170,690 size 136x22; Text 'NumberStyle_2'
   Clock "SecondNeedleHeight" at 330,538 size 150x150
   TextField "Label_SecondNeedleHeight" at 330,690 size 179x22; Text 'SecondNeedleHeight'
   Clock "SecondNeedleWidth" at 490,538 size 150x150
   TextField "Label_SecondNeedleWidth" at 490,690 size 173x22; Text 'SecondNeedleWidth'
   Clock "ShowTicks" at 650,538 size 150x150
   TextField "Label_ShowTicks" at 650,690 size 94x22; Text 'ShowTicks'
   Clock "TickDistance" at 810,538 size 150x150
   TextField "Label_TickDistance" at 810,690 size 113x22; Text 'TickDistance'
   Clock "TickStyle" at 970,538 size 150x150
   TextField "Label_TickStyle" at 970,690 size 84x22; Text 'TickStyle'
   Button "Next" at 1238,776 size 40x22; TextOff 'Text'
      on Click: ActivateScreen("P_Clock_2", 0)

screen "P_Clock_2" 1280x800
   Clock "TicksColor" at 10,10 size 150x150
   TextField "Label_TicksColor" at 10,162 size 94x22; Text 'TicksColor'
   Clock "UseDesignColorSchema" at 170,10 size 150x150
   TextField "Label_UseDesignColorSchema" at 170,162 size 202x22; Text 'UseDesignColorSchema'
   Button "Next" at 1238,776 size 40x22; TextOff 'Text'
      on Click: ActivateScreen("P_Line_1", 0)

